C01873=-23.050,-43.100,93.800,0.0000,0.0000,-150.0000
C01874=-23.050,-38.100,93.800,0.0000,0.0000,-150.0000
C01875=-23.050,-33.100,93.800,0.0000,0.0000,-150.0000
C01876=-23.050,-28.100,93.800,0.0000,0.0000,-150.0000
C01877=-23.050,-23.100,93.800,0.0000,0.0000,-150.0000
C01878=-23.050,-18.100,93.800,0.0000,0.0000,-150.0000
C01879=-23.050,-13.100,93.800,0.0000,0.0000,-150.0000
C01880=-23.050,-8.100,93.800,0.0000,0.0000,-150.0000
C01881=-23.050,-3.100,93.800,0.0000,0.0000,-150.0000
C01882=-23.050,1.900,93.800,0.0000,0.0000,-150.0000
C01883=-23.050,6.900,93.800,0.0000,0.0000,-150.0000
C01884=-23.050,11.900,93.800,0.0000,0.0000,-150.0000
C01885=-23.050,16.900,93.800,0.0000,0.0000,-150.0000
C01886=-23.050,21.900,93.800,0.0000,0.0000,-150.0000
C01887=-23.050,26.900,93.800,0.0000,0.0000,-150.0000
C01888=-23.050,31.900,93.800,0.0000,0.0000,-150.0000
C01889=-23.050,36.900,93.800,0.0000,0.0000,-150.0000
C01890=-23.050,41.900,93.800,0.0000,0.0000,-150.0000
C01891=-18.267,41.900,93.800,0.0000,0.0000,-150.0000
C01892=-13.483,41.900,93.800,0.0000,0.0000,-150.0000
C01893=-8.700,41.900,93.800,0.0000,0.0000,-150.0000
C01894=-3.917,41.900,93.800,0.0000,0.0000,-150.0000
C01895=0.867,41.900,93.800,0.0000,0.0000,-150.0000
C01896=5.650,41.900,93.800,0.0000,0.0000,-150.0000
C01897=10.433,41.900,93.800,0.0000,0.0000,-150.0000
C01898=15.217,41.900,93.800,0.0000,0.0000,-150.0000
C01899=20.000,41.900,93.800,0.0000,0.0000,-150.0000
C01900=25.000,41.900,93.800,0.0000,0.0000,-150.0000
C01901=26.950,43.850,93.800,0.0000,0.0000,-150.0000
C01902=25.000,45.800,93.800,0.0000,0.0000,-150.0000
C01903=20.000,45.800,93.800,0.0000,0.0000,-150.0000
C01904=15.000,45.800,93.800,0.0000,0.0000,-150.0000
C01905=10.000,45.800,93.800,0.0000,0.0000,-150.0000
C01906=5.000,45.800,93.800,0.0000,0.0000,-150.0000
C01907=0.000,45.800,93.800,0.0000,0.0000,-150.0000
C01908=-5.000,45.800,93.800,0.0000,0.0000,-150.0000
C01909=-10.000,45.800,93.800,0.0000,0.0000,-150.0000
C01910=-15.000,45.800,93.800,0.0000,0.0000,-150.0000
C01911=-20.000,45.800,93.800,0.0000,0.0000,-150.0000
C01912=-25.000,45.800,93.800,0.0000,0.0000,-150.0000
C01913=-30.000,45.800,93.800,0.0000,0.0000,-150.0000
C01914=-35.000,45.800,93.800,0.0000,0.0000,-150.0000
C01915=-40.000,45.800,93.800,0.0000,0.0000,-150.0000
C01916=-45.000,45.800,93.800,0.0000,0.0000,-150.0000
C01917=-50.000,45.800,93.800,0.0000,0.0000,-150.0000
C01918=-55.000,45.800,93.800,0.0000,0.0000,-150.0000
C01919=-60.000,45.800,93.800,0.0000,0.0000,-150.0000
C01920=-65.000,45.800,93.800,0.0000,0.0000,-150.0000
C01921=-70.000,45.800,93.800,0.0000,0.0000,-150.0000
C01922=-75.000,45.800,93.800,0.0000,0.0000,-150.0000
C01923=-76.950,43.850,93.800,0.0000,0.0000,-150.0000
C01924=-75.000,41.900,93.800,0.0000,0.0000,-150.0000
C01925=-70.195,41.900,93.800,0.0000,0.0000,-150.0000
C01926=-65.390,41.900,93.800,0.0000,0.0000,-150.0000
C01927=-60.585,41.900,93.800,0.0000,0.0000,-150.0000
C01928=-55.780,41.900,93.800,0.0000,0.0000,-150.0000
C01929=-50.975,41.900,93.800,0.0000,0.0000,-150.0000
C01930=-46.170,41.900,93.800,0.0000,0.0000,-150.0000
C01931=-41.365,41.900,93.800,0.0000,0.0000,-150.0000
C01932=-36.560,41.900,93.800,0.0000,0.0000,-150.0000
C01933=-31.755,41.900,93.800,0.0000,0.0000,-150.0000
C01934=-26.950,41.900,93.800,0.0000,0.0000,-150.0000
C01935=-26.950,36.900,93.800,0.0000,0.0000,-150.0000
C01936=-26.950,31.900,93.800,0.0000,0.0000,-150.0000
C01937=-26.950,26.900,93.800,0.0000,0.0000,-150.0000
C01938=-26.950,21.900,93.800,0.0000,0.0000,-150.0000
C01939=-26.950,16.900,93.800,0.0000,0.0000,-150.0000
C01940=-26.950,11.900,93.800,0.0000,0.0000,-150.0000
C01941=-26.950,6.900,93.800,0.0000,0.0000,-150.0000
C01942=-26.950,1.900,93.800,0.0000,0.0000,-150.0000
C01943=-26.950,-3.100,93.800,0.0000,0.0000,-150.0000
C01944=-26.950,-8.100,93.800,0.0000,0.0000,-150.0000
C01945=-26.950,-13.100,93.800,0.0000,0.0000,-150.0000
C01946=-26.950,-18.100,93.800,0.0000,0.0000,-150.0000
C01947=-26.950,-23.100,93.800,0.0000,0.0000,-150.0000
C01948=-26.950,-28.100,93.800,0.0000,0.0000,-150.0000
C01949=-26.950,-33.100,93.800,0.0000,0.0000,-150.0000
C01950=-26.950,-38.100,93.800,0.0000,0.0000,-150.0000
C01951=-26.950,-43.100,93.800,0.0000,0.0000,-150.0000
C01952=-26.950,-48.100,93.800,0.0000,0.0000,-150.0000
C01953=-26.950,-53.100,93.800,0.0000,0.0000,-150.0000
C01954=-26.950,-58.100,93.800,0.0000,0.0000,-150.0000
C01955=-26.950,-63.100,93.800,0.0000,0.0000,-150.0000
C01956=-26.950,-68.100,93.800,0.0000,0.0000,-150.0000
C01957=-31.755,-68.100,93.800,0.0000,0.0000,-150.0000
C01958=-36.560,-68.100,93.800,0.0000,0.0000,-150.0000
C01959=-41.365,-68.100,93.800,0.0000,0.0000,-150.0000
C01960=-46.170,-68.100,93.800,0.0000,0.0000,-150.0000
C01961=-50.975,-68.100,93.800,0.0000,0.0000,-150.0000
C01962=-55.780,-68.100,93.800,0.0000,0.0000,-150.0000
C01963=-60.585,-68.100,93.800,0.0000,0.0000,-150.0000
C01964=-65.390,-68.100,93.800,0.0000,0.0000,-150.0000
C01965=-70.195,-68.100,93.800,0.0000,0.0000,-150.0000
C01966=-75.000,-68.100,93.800,0.0000,0.0000,-150.0000
C01967=-75.000,-68.100,95.500,0.0000,0.0000,-150.0000
C01968=-70.195,-68.100,95.500,0.0000,0.0000,-150.0000
C01969=-65.390,-68.100,95.500,0.0000,0.0000,-150.0000
C01970=-60.585,-68.100,95.500,0.0000,0.0000,-150.0000
C01971=-55.780,-68.100,95.500,0.0000,0.0000,-150.0000
C01972=-50.975,-68.100,95.500,0.0000,0.0000,-150.0000
C01973=-46.170,-68.100,95.500,0.0000,0.0000,-150.0000
C01974=-41.365,-68.100,95.500,0.0000,0.0000,-150.0000
C01975=-36.560,-68.100,95.500,0.0000,0.0000,-150.0000
C01976=-31.755,-68.100,95.500,0.0000,0.0000,-150.0000
C01977=-26.950,-68.100,95.500,0.0000,0.0000,-150.0000
C01978=-26.950,-63.100,95.500,0.0000,0.0000,-150.0000
C01979=-26.950,-58.100,95.500,0.0000,0.0000,-150.0000
C01980=-26.950,-53.100,95.500,0.0000,0.0000,-150.0000
C01981=-26.950,-48.100,95.500,0.0000,0.0000,-150.0000
C01982=-26.950,-43.100,95.500,0.0000,0.0000,-150.0000
C01983=-26.950,-38.100,95.500,0.0000,0.0000,-150.0000
C01984=-26.950,-33.100,95.500,0.0000,0.0000,-150.0000
C01985=-26.950,-28.100,95.500,0.0000,0.0000,-150.0000
C01986=-26.950,-23.100,95.500,0.0000,0.0000,-150.0000
C01987=-26.950,-18.100,95.500,0.0000,0.0000,-150.0000
C01988=-26.950,-13.100,95.500,0.0000,0.0000,-150.0000
C01989=-26.950,-8.100,95.500,0.0000,0.0000,-150.0000
C01990=-26.950,-3.100,95.500,0.0000,0.0000,-150.0000
C01991=-26.950,1.900,95.500,0.0000,0.0000,-150.0000
C01992=-26.950,6.900,95.500,0.0000,0.0000,-150.0000
C01993=-26.950,11.900,95.500,0.0000,0.0000,-150.0000
C01994=-26.950,16.900,95.500,0.0000,0.0000,-150.0000
C01995=-26.950,21.900,95.500,0.0000,0.0000,-150.0000
C01996=-26.950,26.900,95.500,0.0000,0.0000,-150.0000
C01997=-26.950,31.900,95.500,0.0000,0.0000,-150.0000
C01998=-26.950,36.900,95.500,0.0000,0.0000,-150.0000
C01999=-26.950,41.900,95.500,0.0000,0.0000,-150.0000
C02000=-31.733,41.900,95.500,0.0000,0.0000,-150.0000
C02001=-36.517,41.900,95.500,0.0000,0.0000,-150.0000
C02002=-41.300,41.900,95.500,0.0000,0.0000,-150.0000
C02003=-46.083,41.900,95.500,0.0000,0.0000,-150.0000
C02004=-50.867,41.900,95.500,0.0000,0.0000,-150.0000
C02005=-55.650,41.900,95.500,0.0000,0.0000,-150.0000
C02006=-60.433,41.900,95.500,0.0000,0.0000,-150.0000
C02007=-65.217,41.900,95.500,0.0000,0.0000,-150.0000
C02008=-70.000,41.900,95.500,0.0000,0.0000,-150.0000
C02009=-75.000,41.900,95.500,0.0000,0.0000,-150.0000
C02010=-76.950,43.850,95.500,0.0000,0.0000,-150.0000
C02011=-75.000,45.800,95.500,0.0000,0.0000,-150.0000
C02012=-70.000,45.800,95.500,0.0000,0.0000,-150.0000
C02013=-65.000,45.800,95.500,0.0000,0.0000,-150.0000
C02014=-60.000,45.800,95.500,0.0000,0.0000,-150.0000
C02015=-55.000,45.800,95.500,0.0000,0.0000,-150.0000
C02016=-50.000,45.800,95.500,0.0000,0.0000,-150.0000
C02017=-45.000,45.800,95.500,0.0000,0.0000,-150.0000
C02018=-40.000,45.800,95.500,0.0000,0.0000,-150.0000
C02019=-35.000,45.800,95.500,0.0000,0.0000,-150.0000
C02020=-30.000,45.800,95.500,0.0000,0.0000,-150.0000
C02021=-25.000,45.800,95.500,0.0000,0.0000,-150.0000
C02022=-20.000,45.800,95.500,0.0000,0.0000,-150.0000
C02023=-15.000,45.800,95.500,0.0000,0.0000,-150.0000
C02024=-10.000,45.800,95.500,0.0000,0.0000,-150.0000
C02025=-5.000,45.800,95.500,0.0000,0.0000,-150.0000
C02026=0.000,45.800,95.500,0.0000,0.0000,-150.0000
C02027=5.000,45.800,95.500,0.0000,0.0000,-150.0000
C02028=10.000,45.800,95.500,0.0000,0.0000,-150.0000
C02029=15.000,45.800,95.500,0.0000,0.0000,-150.0000
C02030=20.000,45.800,95.500,0.0000,0.0000,-150.0000
C02031=25.000,45.800,95.500,0.0000,0.0000,-150.0000
C02032=26.950,43.850,95.500,0.0000,0.0000,-150.0000
C02033=25.000,41.900,95.500,0.0000,0.0000,-150.0000
C02034=20.195,41.900,95.500,0.0000,0.0000,-150.0000
C02035=15.390,41.900,95.500,0.0000,0.0000,-150.0000
C02036=10.585,41.900,95.500,0.0000,0.0000,-150.0000
C02037=5.780,41.900,95.500,0.0000,0.0000,-150.0000
C02038=0.975,41.900,95.500,0.0000,0.0000,-150.0000
C02039=-3.830,41.900,95.500,0.0000,0.0000,-150.0000
C02040=-8.635,41.900,95.500,0.0000,0.0000,-150.0000
C02041=-13.440,41.900,95.500,0.0000,0.0000,-150.0000
C02042=-18.245,41.900,95.500,0.0000,0.0000,-150.0000
C02043=-23.050,41.900,95.500,0.0000,0.0000,-150.0000
C02044=-23.050,36.900,95.500,0.0000,0.0000,-150.0000
C02045=-23.050,31.900,95.500,0.0000,0.0000,-150.0000
C02046=-23.050,26.900,95.500,0.0000,0.0000,-150.0000
C02047=-23.050,21.900,95.500,0.0000,0.0000,-150.0000
C02048=-23.050,16.900,95.500,0.0000,0.0000,-150.0000
C02049=-23.050,11.900,95.500,0.0000,0.0000,-150.0000
C02050=-23.050,6.900,95.500,0.0000,0.0000,-150.0000
C02051=-23.050,1.900,95.500,0.0000,0.0000,-150.0000
C02052=-23.050,-3.100,95.500,0.0000,0.0000,-150.0000
C02053=-23.050,-8.100,95.500,0.0000,0.0000,-150.0000
C02054=-23.050,-13.100,95.500,0.0000,0.0000,-150.0000
C02055=-23.050,-18.100,95.500,0.0000,0.0000,-150.0000
C02056=-23.050,-23.100,95.500,0.0000,0.0000,-150.0000
C02057=-23.050,-28.100,95.500,0.0000,0.0000,-150.0000
C02058=-23.050,-33.100,95.500,0.0000,0.0000,-150.0000
C02059=-23.050,-38.100,95.500,0.0000,0.0000,-150.0000
C02060=-23.050,-43.100,95.500,0.0000,0.0000,-150.0000
C02061=-23.050,-48.100,95.500,0.0000,0.0000,-150.0000
C02062=-23.050,-53.100,95.500,0.0000,0.0000,-150.0000
C02063=-23.050,-58.100,95.500,0.0000,0.0000,-150.0000
C02064=-23.050,-63.100,95.500,0.0000,0.0000,-150.0000
C02065=-23.050,-68.100,95.500,0.0000,0.0000,-150.0000
C02066=-18.267,-68.100,95.500,0.0000,0.0000,-150.0000
C02067=-13.483,-68.100,95.500,0.0000,0.0000,-150.0000
C02068=-8.700,-68.100,95.500,0.0000,0.0000,-150.0000
C02069=-3.917,-68.100,95.500,0.0000,0.0000,-150.0000
C02070=0.867,-68.100,95.500,0.0000,0.0000,-150.0000
C02071=5.650,-68.100,95.500,0.0000,0.0000,-150.0000
C02072=10.433,-68.100,95.500,0.0000,0.0000,-150.0000
C02073=15.217,-68.100,95.500,0.0000,0.0000,-150.0000
C02074=20.000,-68.100,95.500,0.0000,0.0000,-150.0000
C02075=25.000,-68.100,95.500,0.0000,0.0000,-150.0000
C02076=26.950,-70.050,95.500,0.0000,0.0000,-150.0000
C02077=25.000,-72.000,95.500,0.0000,0.0000,-150.0000
C02078=20.000,-72.000,95.500,0.0000,0.0000,-150.0000
C02079=15.000,-72.000,95.500,0.0000,0.0000,-150.0000
C02080=10.000,-72.000,95.500,0.0000,0.0000,-150.0000
C02081=5.000,-72.000,95.500,0.0000,0.0000,-150.0000
C02082=0.000,-72.000,95.500,0.0000,0.0000,-150.0000
C02083=-5.000,-72.000,95.500,0.0000,0.0000,-150.0000
C02084=-10.000,-72.000,95.500,0.0000,0.0000,-150.0000
C02085=-15.000,-72.000,95.500,0.0000,0.0000,-150.0000
C02086=-20.000,-72.000,95.500,0.0000,0.0000,-150.0000
C02087=-25.000,-72.000,95.500,0.0000,0.0000,-150.0000
C02088=-30.000,-72.000,95.500,0.0000,0.0000,-150.0000
C02089=-35.000,-72.000,95.500,0.0000,0.0000,-150.0000
C02090=-40.000,-72.000,95.500,0.0000,0.0000,-150.0000
C02091=-45.000,-72.000,95.500,0.0000,0.0000,-150.0000
C02092=-50.000,-72.000,95.500,0.0000,0.0000,-150.0000
C02093=-55.000,-72.000,95.500,0.0000,0.0000,-150.0000
C02094=-60.000,-72.000,95.500,0.0000,0.0000,-150.0000
C02095=-65.000,-72.000,95.500,0.0000,0.0000,-150.0000
C02096=-70.000,-72.000,95.500,0.0000,0.0000,-150.0000
C02097=-75.000,-72.000,95.500,0.0000,0.0000,-150.0000
C02098=-75.000,-72.000,97.200,0.0000,0.0000,-150.0000
C02099=-70.000,-72.000,97.200,0.0000,0.0000,-150.0000
C02100=-65.000,-72.000,97.200,0.0000,0.0000,-150.0000
C02101=-60.000,-72.000,97.200,0.0000,0.0000,-150.0000
C02102=-55.000,-72.000,97.200,0.0000,0.0000,-150.0000
C02103=-50.000,-72.000,97.200,0.0000,0.0000,-150.0000
C02104=-45.000,-72.000,97.200,0.0000,0.0000,-150.0000
C02105=-40.000,-72.000,97.200,0.0000,0.0000,-150.0000
C02106=-35.000,-72.000,97.200,0.0000,0.0000,-150.0000
C02107=-30.000,-72.000,97.200,0.0000,0.0000,-150.0000
C02108=-25.000,-72.000,97.200,0.0000,0.0000,-150.0000
C02109=-20.000,-72.000,97.200,0.0000,0.0000,-150.0000
C02110=-15.000,-72.000,97.200,0.0000,0.0000,-150.0000
C02111=-10.000,-72.000,97.200,0.0000,0.0000,-150.0000
C02112=-5.000,-72.000,97.200,0.0000,0.0000,-150.0000
C02113=0.000,-72.000,97.200,0.0000,0.0000,-150.0000
C02114=5.000,-72.000,97.200,0.0000,0.0000,-150.0000
C02115=10.000,-72.000,97.200,0.0000,0.0000,-150.0000
C02116=15.000,-72.000,97.200,0.0000,0.0000,-150.0000
C02117=20.000,-72.000,97.200,0.0000,0.0000,-150.0000
C02118=25.000,-72.000,97.200,0.0000,0.0000,-150.0000
C02119=26.950,-70.050,97.200,0.0000,0.0000,-150.0000
C02120=25.000,-68.100,97.200,0.0000,0.0000,-150.0000
C02121=20.195,-68.100,97.200,0.0000,0.0000,-150.0000
C02122=15.390,-68.100,97.200,0.0000,0.0000,-150.0000
C02123=10.585,-68.100,97.200,0.0000,0.0000,-150.0000
C02124=5.780,-68.100,97.200,0.0000,0.0000,-150.0000
C02125=0.975,-68.100,97.200,0.0000,0.0000,-150.0000
C02126=-3.830,-68.100,97.200,0.0000,0.0000,-150.0000
C02127=-8.635,-68.100,97.200,0.0000,0.0000,-150.0000
C02128=-13.440,-68.100,97.200,0.0000,0.0000,-150.0000
C02129=-18.245,-68.100,97.200,0.0000,0.0000,-150.0000
C02130=-23.050,-68.100,97.200,0.0000,0.0000,-150.0000
C02131=-23.050,-63.100,97.200,0.0000,0.0000,-150.0000
C02132=-23.050,-58.100,97.200,0.0000,0.0000,-150.0000
C02133=-23.050,-53.100,97.200,0.0000,0.0000,-150.0000
C02134=-23.050,-48.100,97.200,0.0000,0.0000,-150.0000
C02135=-23.050,-43.100,97.200,0.0000,0.0000,-150.0000
C02136=-23.050,-38.100,97.200,0.0000,0.0000,-150.0000
C02137=-23.050,-33.100,97.200,0.0000,0.0000,-150.0000
C02138=-23.050,-28.100,97.200,0.0000,0.0000,-150.0000
C02139=-23.050,-23.100,97.200,0.0000,0.0000,-150.0000
C02140=-23.050,-18.100,97.200,0.0000,0.0000,-150.0000
C02141=-23.050,-13.100,97.200,0.0000,0.0000,-150.0000
C02142=-23.050,-8.100,97.200,0.0000,0.0000,-150.0000
C02143=-23.050,-3.100,97.200,0.0000,0.0000,-150.0000
C02144=-23.050,1.900,97.200,0.0000,0.0000,-150.0000
C02145=-23.050,6.900,97.200,0.0000,0.0000,-150.0000
C02146=-23.050,11.900,97.200,0.0000,0.0000,-150.0000
C02147=-23.050,16.900,97.200,0.0000,0.0000,-150.0000
C02148=-23.050,21.900,97.200,0.0000,0.0000,-150.0000
C02149=-23.050,26.900,97.200,0.0000,0.0000,-150.0000
C02150=-23.050,31.900,97.200,0.0000,0.0000,-150.0000
C02151=-23.050,36.900,97.200,0.0000,0.0000,-150.0000
C02152=-23.050,41.900,97.200,0.0000,0.0000,-150.0000
C02153=-18.267,41.900,97.200,0.0000,0.0000,-150.0000
C02154=-13.483,41.900,97.200,0.0000,0.0000,-150.0000
C02155=-8.700,41.900,97.200,0.0000,0.0000,-150.0000
C02156=-3.917,41.900,97.200,0.0000,0.0000,-150.0000
C02157=0.867,41.900,97.200,0.0000,0.0000,-150.0000
C02158=5.650,41.900,97.200,0.0000,0.0000,-150.0000
C02159=10.433,41.900,97.200,0.0000,0.0000,-150.0000
C02160=15.217,41.900,97.200,0.0000,0.0000,-150.0000
C02161=20.000,41.900,97.200,0.0000,0.0000,-150.0000
C02162=25.000,41.900,97.200,0.0000,0.0000,-150.0000
C02163=26.950,43.850,97.200,0.0000,0.0000,-150.0000
C02164=25.000,45.800,97.200,0.0000,0.0000,-150.0000
C02165=20.000,45.800,97.200,0.0000,0.0000,-150.0000
C02166=15.000,45.800,97.200,0.0000,0.0000,-150.0000
C02167=10.000,45.800,97.200,0.0000,0.0000,-150.0000
C02168=5.000,45.800,97.200,0.0000,0.0000,-150.0000
C02169=0.000,45.800,97.200,0.0000,0.0000,-150.0000
C02170=-5.000,45.800,97.200,0.0000,0.0000,-150.0000
C02171=-10.000,45.800,97.200,0.0000,0.0000,-150.0000
C02172=-15.000,45.800,97.200,0.0000,0.0000,-150.0000
C02173=-20.000,45.800,97.200,0.0000,0.0000,-150.0000
C02174=-25.000,45.800,97.200,0.0000,0.0000,-150.0000
C02175=-30.000,45.800,97.200,0.0000,0.0000,-150.0000
C02176=-35.000,45.800,97.200,0.0000,0.0000,-150.0000
C02177=-40.000,45.800,97.200,0.0000,0.0000,-150.0000
C02178=-45.000,45.800,97.200,0.0000,0.0000,-150.0000
C02179=-50.000,45.800,97.200,0.0000,0.0000,-150.0000
C02180=-55.000,45.800,97.200,0.0000,0.0000,-150.0000
C02181=-60.000,45.800,97.200,0.0000,0.0000,-150.0000
C02182=-65.000,45.800,97.200,0.0000,0.0000,-150.0000
C02183=-70.000,45.800,97.200,0.0000,0.0000,-150.0000
C02184=-75.000,45.800,97.200,0.0000,0.0000,-150.0000
C02185=-76.950,43.850,97.200,0.0000,0.0000,-150.0000
C02186=-75.000,41.900,97.200,0.0000,0.0000,-150.0000
C02187=-70.195,41.900,97.200,0.0000,0.0000,-150.0000
C02188=-65.390,41.900,97.200,0.0000,0.0000,-150.0000
C02189=-60.585,41.900,97.200,0.0000,0.0000,-150.0000
C02190=-55.780,41.900,97.200,0.0000,0.0000,-150.0000
C02191=-50.975,41.900,97.200,0.0000,0.0000,-150.0000
C02192=-46.170,41.900,97.200,0.0000,0.0000,-150.0000
C02193=-41.365,41.900,97.200,0.0000,0.0000,-150.0000
C02194=-36.560,41.900,97.200,0.0000,0.0000,-150.0000
C02195=-31.755,41.900,97.200,0.0000,0.0000,-150.0000
C02196=-26.950,41.900,97.200,0.0000,0.0000,-150.0000
C02197=-26.950,36.900,97.200,0.0000,0.0000,-150.0000
C02198=-26.950,31.900,97.200,0.0000,0.0000,-150.0000
C02199=-26.950,26.900,97.200,0.0000,0.0000,-150.0000
C02200=-26.950,21.900,97.200,0.0000,0.0000,-150.0000
C02201=-26.950,16.900,97.200,0.0000,0.0000,-150.0000
C02202=-26.950,11.900,97.200,0.0000,0.0000,-150.0000
C02203=-26.950,6.900,97.200,0.0000,0.0000,-150.0000
C02204=-26.950,1.900,97.200,0.0000,0.0000,-150.0000
C02205=-26.950,-3.100,97.200,0.0000,0.0000,-150.0000
C02206=-26.950,-8.100,97.200,0.0000,0.0000,-150.0000
C02207=-26.950,-13.100,97.200,0.0000,0.0000,-150.0000
C02208=-26.950,-18.100,97.200,0.0000,0.0000,-150.0000
C02209=-26.950,-23.100,97.200,0.0000,0.0000,-150.0000
C02210=-26.950,-28.100,97.200,0.0000,0.0000,-150.0000
C02211=-26.950,-33.100,97.200,0.0000,0.0000,-150.0000
C02212=-26.950,-38.100,97.200,0.0000,0.0000,-150.0000
C02213=-26.950,-43.100,97.200,0.0000,0.0000,-150.0000
C02214=-26.950,-48.100,97.200,0.0000,0.0000,-150.0000
C02215=-26.950,-53.100,97.200,0.0000,0.0000,-150.0000
C02216=-26.950,-58.100,97.200,0.0000,0.0000,-150.0000
C02217=-26.950,-63.100,97.200,0.0000,0.0000,-150.0000
C02218=-26.950,-68.100,97.200,0.0000,0.0000,-150.0000
C02219=-31.755,-68.100,97.200,0.0000,0.0000,-150.0000
C02220=-36.560,-68.100,97.200,0.0000,0.0000,-150.0000
C02221=-41.365,-68.100,97.200,0.0000,0.0000,-150.0000
C02222=-46.170,-68.100,97.200,0.0000,0.0000,-150.0000
C02223=-50.975,-68.100,97.200,0.0000,0.0000,-150.0000
C02224=-55.780,-68.100,97.200,0.0000,0.0000,-150.0000
C02225=-60.585,-68.100,97.200,0.0000,0.0000,-150.0000
C02226=-65.390,-68.100,97.200,0.0000,0.0000,-150.0000
C02227=-70.195,-68.100,97.200,0.0000,0.0000,-150.0000
C02228=-75.000,-68.100,97.200,0.0000,0.0000,-150.0000
C02229=-75.000,-68.100,98.900,0.0000,0.0000,-150.0000
C02230=-70.195,-68.100,98.900,0.0000,0.0000,-150.0000
C02231=-65.390,-68.100,98.900,0.0000,0.0000,-150.0000
C02232=-60.585,-68.100,98.900,0.0000,0.0000,-150.0000
C02233=-55.780,-68.100,98.900,0.0000,0.0000,-150.0000
C02234=-50.975,-68.100,98.900,0.0000,0.0000,-150.0000
C02235=-46.170,-68.100,98.900,0.0000,0.0000,-150.0000
C02236=-41.365,-68.100,98.900,0.0000,0.0000,-150.0000
C02237=-36.560,-68.100,98.900,0.0000,0.0000,-150.0000
C02238=-31.755,-68.100,98.900,0.0000,0.0000,-150.0000
C02239=-26.950,-68.100,98.900,0.0000,0.0000,-150.0000
C02240=-26.950,-63.100,98.900,0.0000,0.0000,-150.0000
C02241=-26.950,-58.100,98.900,0.0000,0.0000,-150.0000
C02242=-26.950,-53.100,98.900,0.0000,0.0000,-150.0000
C02243=-26.950,-48.100,98.900,0.0000,0.0000,-150.0000
C02244=-26.950,-43.100,98.900,0.0000,0.0000,-150.0000
C02245=-26.950,-38.100,98.900,0.0000,0.0000,-150.0000
C02246=-26.950,-33.100,98.900,0.0000,0.0000,-150.0000
C02247=-26.950,-28.100,98.900,0.0000,0.0000,-150.0000
C02248=-26.950,-23.100,98.900,0.0000,0.0000,-150.0000
C02249=-26.950,-18.100,98.900,0.0000,0.0000,-150.0000
C02250=-26.950,-13.100,98.900,0.0000,0.0000,-150.0000
C02251=-26.950,-8.100,98.900,0.0000,0.0000,-150.0000
C02252=-26.950,-3.100,98.900,0.0000,0.0000,-150.0000
C02253=-26.950,1.900,98.900,0.0000,0.0000,-150.0000
C02254=-26.950,6.900,98.900,0.0000,0.0000,-150.0000
C02255=-26.950,11.900,98.900,0.0000,0.0000,-150.0000
C02256=-26.950,16.900,98.900,0.0000,0.0000,-150.0000
C02257=-26.950,21.900,98.900,0.0000,0.0000,-150.0000
C02258=-26.950,26.900,98.900,0.0000,0.0000,-150.0000
C02259=-26.950,31.900,98.900,0.0000,0.0000,-150.0000
C02260=-26.950,36.900,98.900,0.0000,0.0000,-150.0000
C02261=-26.950,41.900,98.900,0.0000,0.0000,-150.0000
C02262=-31.733,41.900,98.900,0.0000,0.0000,-150.0000
C02263=-36.517,41.900,98.900,0.0000,0.0000,-150.0000
C02264=-41.300,41.900,98.900,0.0000,0.0000,-150.0000
C02265=-46.083,41.900,98.900,0.0000,0.0000,-150.0000
C02266=-50.867,41.900,98.900,0.0000,0.0000,-150.0000
C02267=-55.650,41.900,98.900,0.0000,0.0000,-150.0000
C02268=-60.433,41.900,98.900,0.0000,0.0000,-150.0000
C02269=-65.217,41.900,98.900,0.0000,0.0000,-150.0000
C02270=-70.000,41.900,98.900,0.0000,0.0000,-150.0000
C02271=-75.000,41.900,98.900,0.0000,0.0000,-150.0000
C02272=-76.950,43.850,98.900,0.0000,0.0000,-150.0000
C02273=-75.000,45.800,98.900,0.0000,0.0000,-150.0000
C02274=-70.000,45.800,98.900,0.0000,0.0000,-150.0000
C02275=-65.000,45.800,98.900,0.0000,0.0000,-150.0000
C02276=-60.000,45.800,98.900,0.0000,0.0000,-150.0000
C02277=-55.000,45.800,98.900,0.0000,0.0000,-150.0000
C02278=-50.000,45.800,98.900,0.0000,0.0000,-150.0000
C02279=-45.000,45.800,98.900,0.0000,0.0000,-150.0000
C02280=-40.000,45.800,98.900,0.0000,0.0000,-150.0000
C02281=-35.000,45.800,98.900,0.0000,0.0000,-150.0000
C02282=-30.000,45.800,98.900,0.0000,0.0000,-150.0000
C02283=-25.000,45.800,98.900,0.0000,0.0000,-150.0000
C02284=-20.000,45.800,98.900,0.0000,0.0000,-150.0000
C02285=-15.000,45.800,98.900,0.0000,0.0000,-150.0000
C02286=-10.000,45.800,98.900,0.0000,0.0000,-150.0000
C02287=-5.000,45.800,98.900,0.0000,0.0000,-150.0000
C02288=0.000,45.800,98.900,0.0000,0.0000,-150.0000
C02289=5.000,45.800,98.900,0.0000,0.0000,-150.0000
C02290=10.000,45.800,98.900,0.0000,0.0000,-150.0000
C02291=15.000,45.800,98.900,0.0000,0.0000,-150.0000
C02292=20.000,45.800,98.900,0.0000,0.0000,-150.0000
C02293=25.000,45.800,98.900,0.0000,0.0000,-150.0000
C02294=26.950,43.850,98.900,0.0000,0.0000,-150.0000
C02295=25.000,41.900,98.900,0.0000,0.0000,-150.0000
C02296=20.195,41.900,98.900,0.0000,0.0000,-150.0000
C02297=15.390,41.900,98.900,0.0000,0.0000,-150.0000
C02298=10.585,41.900,98.900,0.0000,0.0000,-150.0000
C02299=5.780,41.900,98.900,0.0000,0.0000,-150.0000
C02300=0.975,41.900,98.900,0.0000,0.0000,-150.0000
C02301=-3.830,41.900,98.900,0.0000,0.0000,-150.0000
C02302=-8.635,41.900,98.900,0.0000,0.0000,-150.0000
C02303=-13.440,41.900,98.900,0.0000,0.0000,-150.0000
C02304=-18.245,41.900,98.900,0.0000,0.0000,-150.0000
C02305=-23.050,41.900,98.900,0.0000,0.0000,-150.0000
C02306=-23.050,36.900,98.900,0.0000,0.0000,-150.0000
C02307=-23.050,31.900,98.900,0.0000,0.0000,-150.0000
C02308=-23.050,26.900,98.900,0.0000,0.0000,-150.0000
C02309=-23.050,21.900,98.900,0.0000,0.0000,-150.0000
C02310=-23.050,16.900,98.900,0.0000,0.0000,-150.0000
C02311=-23.050,11.900,98.900,0.0000,0.0000,-150.0000
C02312=-23.050,6.900,98.900,0.0000,0.0000,-150.0000
C02313=-23.050,1.900,98.900,0.0000,0.0000,-150.0000
C02314=-23.050,-3.100,98.900,0.0000,0.0000,-150.0000
C02315=-23.050,-8.100,98.900,0.0000,0.0000,-150.0000
C02316=-23.050,-13.100,98.900,0.0000,0.0000,-150.0000
C02317=-23.050,-18.100,98.900,0.0000,0.0000,-150.0000
C02318=-23.050,-23.100,98.900,0.0000,0.0000,-150.0000
C02319=-23.050,-28.100,98.900,0.0000,0.0000,-150.0000
C02320=-23.050,-33.100,98.900,0.0000,0.0000,-150.0000
C02321=-23.050,-38.100,98.900,0.0000,0.0000,-150.0000
C02322=-23.050,-43.100,98.900,0.0000,0.0000,-150.0000
C02323=-23.050,-48.100,98.900,0.0000,0.0000,-150.0000
C02324=-23.050,-53.100,98.900,0.0000,0.0000,-150.0000
C02325=-23.050,-58.100,98.900,0.0000,0.0000,-150.0000
C02326=-23.050,-63.100,98.900,0.0000,0.0000,-150.0000
C02327=-23.050,-68.100,98.900,0.0000,0.0000,-150.0000
C02328=-18.267,-68.100,98.900,0.0000,0.0000,-150.0000
C02329=-13.483,-68.100,98.900,0.0000,0.0000,-150.0000
C02330=-8.700,-68.100,98.900,0.0000,0.0000,-150.0000
C02331=-3.917,-68.100,98.900,0.0000,0.0000,-150.0000
C02332=0.867,-68.100,98.900,0.0000,0.0000,-150.0000
C02333=5.650,-68.100,98.900,0.0000,0.0000,-150.0000
C02334=10.433,-68.100,98.900,0.0000,0.0000,-150.0000
C02335=15.217,-68.100,98.900,0.0000,0.0000,-150.0000
C02336=20.000,-68.100,98.900,0.0000,0.0000,-150.0000
C02337=25.000,-68.100,98.900,0.0000,0.0000,-150.0000
C02338=26.950,-70.050,98.900,0.0000,0.0000,-150.0000
C02339=25.000,-72.000,98.900,0.0000,0.0000,-150.0000
C02340=20.000,-72.000,98.900,0.0000,0.0000,-150.0000
C02341=15.000,-72.000,98.900,0.0000,0.0000,-150.0000
C02342=10.000,-72.000,98.900,0.0000,0.0000,-150.0000
C02343=5.000,-72.000,98.900,0.0000,0.0000,-150.0000
C02344=0.000,-72.000,98.900,0.0000,0.0000,-150.0000
C02345=-5.000,-72.000,98.900,0.0000,0.0000,-150.0000
C02346=-10.000,-72.000,98.900,0.0000,0.0000,-150.0000
C02347=-15.000,-72.000,98.900,0.0000,0.0000,-150.0000
C02348=-20.000,-72.000,98.900,0.0000,0.0000,-150.0000
C02349=-25.000,-72.000,98.900,0.0000,0.0000,-150.0000
C02350=-30.000,-72.000,98.900,0.0000,0.0000,-150.0000
C02351=-35.000,-72.000,98.900,0.0000,0.0000,-150.0000
C02352=-40.000,-72.000,98.900,0.0000,0.0000,-150.0000
C02353=-45.000,-72.000,98.900,0.0000,0.0000,-150.0000
C02354=-50.000,-72.000,98.900,0.0000,0.0000,-150.0000
C02355=-55.000,-72.000,98.900,0.0000,0.0000,-150.0000
C02356=-60.000,-72.000,98.900,0.0000,0.0000,-150.0000
C02357=-65.000,-72.000,98.900,0.0000,0.0000,-150.0000
C02358=-70.000,-72.000,98.900,0.0000,0.0000,-150.0000
C02359=-75.000,-72.000,98.900,0.0000,0.0000,-150.0000
C02360=-75.000,-72.000,100.600,0.0000,0.0000,-150.0000
C02361=-70.000,-72.000,100.600,0.0000,0.0000,-150.0000
C02362=-65.000,-72.000,100.600,0.0000,0.0000,-150.0000
C02363=-60.000,-72.000,100.600,0.0000,0.0000,-150.0000
C02364=-55.000,-72.000,100.600,0.0000,0.0000,-150.0000
C02365=-50.000,-72.000,100.600,0.0000,0.0000,-150.0000
C02366=-45.000,-72.000,100.600,0.0000,0.0000,-150.0000
C02367=-40.000,-72.000,100.600,0.0000,0.0000,-150.0000
C02368=-35.000,-72.000,100.600,0.0000,0.0000,-150.0000
C02369=-30.000,-72.000,100.600,0.0000,0.0000,-150.0000
C02370=-25.000,-72.000,100.600,0.0000,0.0000,-150.0000
C02371=-20.000,-72.000,100.600,0.0000,0.0000,-150.0000
C02372=-15.000,-72.000,100.600,0.0000,0.0000,-150.0000
C02373=-10.000,-72.000,100.600,0.0000,0.0000,-150.0000
C02374=-5.000,-72.000,100.600,0.0000,0.0000,-150.0000
C02375=0.000,-72.000,100.600,0.0000,0.0000,-150.0000
C02376=5.000,-72.000,100.600,0.0000,0.0000,-150.0000
C02377=10.000,-72.000,100.600,0.0000,0.0000,-150.0000
C02378=15.000,-72.000,100.600,0.0000,0.0000,-150.0000
C02379=20.000,-72.000,100.600,0.0000,0.0000,-150.0000
C02380=25.000,-72.000,100.600,0.0000,0.0000,-150.0000
C02381=26.950,-70.050,100.600,0.0000,0.0000,-150.0000
C02382=25.000,-68.100,100.600,0.0000,0.0000,-150.0000
C02383=20.195,-68.100,100.600,0.0000,0.0000,-150.0000
C02384=15.390,-68.100,100.600,0.0000,0.0000,-150.0000
C02385=10.585,-68.100,100.600,0.0000,0.0000,-150.0000
C02386=5.780,-68.100,100.600,0.0000,0.0000,-150.0000
C02387=0.975,-68.100,100.600,0.0000,0.0000,-150.0000
C02388=-3.830,-68.100,100.600,0.0000,0.0000,-150.0000
C02389=-8.635,-68.100,100.600,0.0000,0.0000,-150.0000
C02390=-13.440,-68.100,100.600,0.0000,0.0000,-150.0000
C02391=-18.245,-68.100,100.600,0.0000,0.0000,-150.0000
C02392=-23.050,-68.100,100.600,0.0000,0.0000,-150.0000
C02393=-23.050,-63.100,100.600,0.0000,0.0000,-150.0000
C02394=-23.050,-58.100,100.600,0.0000,0.0000,-150.0000
C02395=-23.050,-53.100,100.600,0.0000,0.0000,-150.0000
C02396=-23.050,-48.100,100.600,0.0000,0.0000,-150.0000
C02397=-23.050,-43.100,100.600,0.0000,0.0000,-150.0000
C02398=-23.050,-38.100,100.600,0.0000,0.0000,-150.0000
C02399=-23.050,-33.100,100.600,0.0000,0.0000,-150.0000
C02400=-23.050,-28.100,100.600,0.0000,0.0000,-150.0000
C02401=-23.050,-23.100,100.600,0.0000,0.0000,-150.0000
C02402=-23.050,-18.100,100.600,0.0000,0.0000,-150.0000
C02403=-23.050,-13.100,100.600,0.0000,0.0000,-150.0000
C02404=-23.050,-8.100,100.600,0.0000,0.0000,-150.0000
C02405=-23.050,-3.100,100.600,0.0000,0.0000,-150.0000
C02406=-23.050,1.900,100.600,0.0000,0.0000,-150.0000
C02407=-23.050,6.900,100.600,0.0000,0.0000,-150.0000
C02408=-23.050,11.900,100.600,0.0000,0.0000,-150.0000
C02409=-23.050,16.900,100.600,0.0000,0.0000,-150.0000
C02410=-23.050,21.900,100.600,0.0000,0.0000,-150.0000
C02411=-23.050,26.900,100.600,0.0000,0.0000,-150.0000
C02412=-23.050,31.900,100.600,0.0000,0.0000,-150.0000
C02413=-23.050,36.900,100.600,0.0000,0.0000,-150.0000
C02414=-23.050,41.900,100.600,0.0000,0.0000,-150.0000
C02415=-18.267,41.900,100.600,0.0000,0.0000,-150.0000
C02416=-13.483,41.900,100.600,0.0000,0.0000,-150.0000
C02417=-8.700,41.900,100.600,0.0000,0.0000,-150.0000
C02418=-3.917,41.900,100.600,0.0000,0.0000,-150.0000
C02419=0.867,41.900,100.600,0.0000,0.0000,-150.0000
C02420=5.650,41.900,100.600,0.0000,0.0000,-150.0000
C02421=10.433,41.900,100.600,0.0000,0.0000,-150.0000
C02422=15.217,41.900,100.600,0.0000,0.0000,-150.0000
C02423=20.000,41.900,100.600,0.0000,0.0000,-150.0000
C02424=25.000,41.900,100.600,0.0000,0.0000,-150.0000
C02425=26.950,43.850,100.600,0.0000,0.0000,-150.0000
C02426=25.000,45.800,100.600,0.0000,0.0000,-150.0000
C02427=20.000,45.800,100.600,0.0000,0.0000,-150.0000
C02428=15.000,45.800,100.600,0.0000,0.0000,-150.0000
C02429=10.000,45.800,100.600,0.0000,0.0000,-150.0000
C02430=5.000,45.800,100.600,0.0000,0.0000,-150.0000
C02431=0.000,45.800,100.600,0.0000,0.0000,-150.0000
C02432=-5.000,45.800,100.600,0.0000,0.0000,-150.0000
C02433=-10.000,45.800,100.600,0.0000,0.0000,-150.0000
C02434=-15.000,45.800,100.600,0.0000,0.0000,-150.0000
C02435=-20.000,45.800,100.600,0.0000,0.0000,-150.0000
C02436=-25.000,45.800,100.600,0.0000,0.0000,-150.0000
C02437=-30.000,45.800,100.600,0.0000,0.0000,-150.0000
C02438=-35.000,45.800,100.600,0.0000,0.0000,-150.0000
C02439=-40.000,45.800,100.600,0.0000,0.0000,-150.0000
C02440=-45.000,45.800,100.600,0.0000,0.0000,-150.0000
C02441=-50.000,45.800,100.600,0.0000,0.0000,-150.0000
C02442=-55.000,45.800,100.600,0.0000,0.0000,-150.0000
C02443=-60.000,45.800,100.600,0.0000,0.0000,-150.0000
C02444=-65.000,45.800,100.600,0.0000,0.0000,-150.0000
C02445=-70.000,45.800,100.600,0.0000,0.0000,-150.0000
C02446=-75.000,45.800,100.600,0.0000,0.0000,-150.0000
C02447=-76.950,43.850,100.600,0.0000,0.0000,-150.0000
C02448=-75.000,41.900,100.600,0.0000,0.0000,-150.0000
C02449=-70.195,41.900,100.600,0.0000,0.0000,-150.0000
C02450=-65.390,41.900,100.600,0.0000,0.0000,-150.0000
C02451=-60.585,41.900,100.600,0.0000,0.0000,-150.0000
C02452=-55.780,41.900,100.600,0.0000,0.0000,-150.0000
C02453=-50.975,41.900,100.600,0.0000,0.0000,-150.0000
C02454=-46.170,41.900,100.600,0.0000,0.0000,-150.0000
C02455=-41.365,41.900,100.600,0.0000,0.0000,-150.0000
C02456=-36.560,41.900,100.600,0.0000,0.0000,-150.0000
C02457=-31.755,41.900,100.600,0.0000,0.0000,-150.0000
C02458=-26.950,41.900,100.600,0.0000,0.0000,-150.0000
C02459=-26.950,36.900,100.600,0.0000,0.0000,-150.0000
C02460=-26.950,31.900,100.600,0.0000,0.0000,-150.0000
C02461=-26.950,26.900,100.600,0.0000,0.0000,-150.0000
C02462=-26.950,21.900,100.600,0.0000,0.0000,-150.0000
C02463=-26.950,16.900,100.600,0.0000,0.0000,-150.0000
C02464=-26.950,11.900,100.600,0.0000,0.0000,-150.0000
C02465=-26.950,6.900,100.600,0.0000,0.0000,-150.0000
C02466=-26.950,1.900,100.600,0.0000,0.0000,-150.0000
C02467=-26.950,-3.100,100.600,0.0000,0.0000,-150.0000
C02468=-26.950,-8.100,100.600,0.0000,0.0000,-150.0000
C02469=-26.950,-13.100,100.600,0.0000,0.0000,-150.0000
C02470=-26.950,-18.100,100.600,0.0000,0.0000,-150.0000
C02471=-26.950,-23.100,100.600,0.0000,0.0000,-150.0000
C02472=-26.950,-28.100,100.600,0.0000,0.0000,-150.0000
C02473=-26.950,-33.100,100.600,0.0000,0.0000,-150.0000
C02474=-26.950,-38.100,100.600,0.0000,0.0000,-150.0000
C02475=-26.950,-43.100,100.600,0.0000,0.0000,-150.0000
C02476=-26.950,-48.100,100.600,0.0000,0.0000,-150.0000
C02477=-26.950,-53.100,100.600,0.0000,0.0000,-150.0000
C02478=-26.950,-58.100,100.600,0.0000,0.0000,-150.0000
C02479=-26.950,-63.100,100.600,0.0000,0.0000,-150.0000
C02480=-26.950,-68.100,100.600,0.0000,0.0000,-150.0000
C02481=-31.755,-68.100,100.600,0.0000,0.0000,-150.0000
C02482=-36.560,-68.100,100.600,0.0000,0.0000,-150.0000
C02483=-41.365,-68.100,100.600,0.0000,0.0000,-150.0000
C02484=-46.170,-68.100,100.600,0.0000,0.0000,-150.0000
C02485=-50.975,-68.100,100.600,0.0000,0.0000,-150.0000
C02486=-55.780,-68.100,100.600,0.0000,0.0000,-150.0000
C02487=-60.585,-68.100,100.600,0.0000,0.0000,-150.0000
C02488=-65.390,-68.100,100.600,0.0000,0.0000,-150.0000
C02489=-70.195,-68.100,100.600,0.0000,0.0000,-150.0000
C02490=-75.000,-68.100,100.600,0.0000,0.0000,-150.0000
C02491=-75.000,-68.100,102.300,0.0000,0.0000,-150.0000
C02492=-70.195,-68.100,102.300,0.0000,0.0000,-150.0000
C02493=-65.390,-68.100,102.300,0.0000,0.0000,-150.0000
C02494=-60.585,-68.100,102.300,0.0000,0.0000,-150.0000
C02495=-55.780,-68.100,102.300,0.0000,0.0000,-150.0000
C02496=-50.975,-68.100,102.300,0.0000,0.0000,-150.0000
C02497=-46.170,-68.100,102.300,0.0000,0.0000,-150.0000
C02498=-41.365,-68.100,102.300,0.0000,0.0000,-150.0000
C02499=-36.560,-68.100,102.300,0.0000,0.0000,-150.0000
C02500=-31.755,-68.100,102.300,0.0000,0.0000,-150.0000
C02501=-26.950,-68.100,102.300,0.0000,0.0000,-150.0000
C02502=-26.950,-63.100,102.300,0.0000,0.0000,-150.0000
C02503=-26.950,-58.100,102.300,0.0000,0.0000,-150.0000
C02504=-26.950,-53.100,102.300,0.0000,0.0000,-150.0000
C02505=-26.950,-48.100,102.300,0.0000,0.0000,-150.0000
C02506=-26.950,-43.100,102.300,0.0000,0.0000,-150.0000
C02507=-26.950,-38.100,102.300,0.0000,0.0000,-150.0000
C02508=-26.950,-33.100,102.300,0.0000,0.0000,-150.0000
C02509=-26.950,-28.100,102.300,0.0000,0.0000,-150.0000
C02510=-26.950,-23.100,102.300,0.0000,0.0000,-150.0000
C02511=-26.950,-18.100,102.300,0.0000,0.0000,-150.0000
C02512=-26.950,-13.100,102.300,0.0000,0.0000,-150.0000
C02513=-26.950,-8.100,102.300,0.0000,0.0000,-150.0000
C02514=-26.950,-3.100,102.300,0.0000,0.0000,-150.0000
C02515=-26.950,1.900,102.300,0.0000,0.0000,-150.0000
C02516=-26.950,6.900,102.300,0.0000,0.0000,-150.0000
C02517=-26.950,11.900,102.300,0.0000,0.0000,-150.0000
C02518=-26.950,16.900,102.300,0.0000,0.0000,-150.0000
C02519=-26.950,21.900,102.300,0.0000,0.0000,-150.0000
C02520=-26.950,26.900,102.300,0.0000,0.0000,-150.0000
C02521=-26.950,31.900,102.300,0.0000,0.0000,-150.0000
C02522=-26.950,36.900,102.300,0.0000,0.0000,-150.0000
C02523=-26.950,41.900,102.300,0.0000,0.0000,-150.0000
C02524=-31.733,41.900,102.300,0.0000,0.0000,-150.0000
C02525=-36.517,41.900,102.300,0.0000,0.0000,-150.0000
C02526=-41.300,41.900,102.300,0.0000,0.0000,-150.0000
C02527=-46.083,41.900,102.300,0.0000,0.0000,-150.0000
C02528=-50.867,41.900,102.300,0.0000,0.0000,-150.0000
C02529=-55.650,41.900,102.300,0.0000,0.0000,-150.0000
C02530=-60.433,41.900,102.300,0.0000,0.0000,-150.0000
C02531=-65.217,41.900,102.300,0.0000,0.0000,-150.0000
C02532=-70.000,41.900,102.300,0.0000,0.0000,-150.0000
C02533=-75.000,41.900,102.300,0.0000,0.0000,-150.0000
C02534=-76.950,43.850,102.300,0.0000,0.0000,-150.0000
C02535=-75.000,45.800,102.300,0.0000,0.0000,-150.0000
C02536=-70.000,45.800,102.300,0.0000,0.0000,-150.0000
C02537=-65.000,45.800,102.300,0.0000,0.0000,-150.0000
C02538=-60.000,45.800,102.300,0.0000,0.0000,-150.0000
C02539=-55.000,45.800,102.300,0.0000,0.0000,-150.0000
C02540=-50.000,45.800,102.300,0.0000,0.0000,-150.0000
C02541=-45.000,45.800,102.300,0.0000,0.0000,-150.0000
C02542=-40.000,45.800,102.300,0.0000,0.0000,-150.0000
C02543=-35.000,45.800,102.300,0.0000,0.0000,-150.0000
C02544=-30.000,45.800,102.300,0.0000,0.0000,-150.0000
C02545=-25.000,45.800,102.300,0.0000,0.0000,-150.0000
C02546=-20.000,45.800,102.300,0.0000,0.0000,-150.0000
C02547=-15.000,45.800,102.300,0.0000,0.0000,-150.0000
C02548=-10.000,45.800,102.300,0.0000,0.0000,-150.0000
C02549=-5.000,45.800,102.300,0.0000,0.0000,-150.0000
C02550=0.000,45.800,102.300,0.0000,0.0000,-150.0000
C02551=5.000,45.800,102.300,0.0000,0.0000,-150.0000
C02552=10.000,45.800,102.300,0.0000,0.0000,-150.0000
C02553=15.000,45.800,102.300,0.0000,0.0000,-150.0000
C02554=20.000,45.800,102.300,0.0000,0.0000,-150.0000
C02555=25.000,45.800,102.300,0.0000,0.0000,-150.0000
C02556=26.950,43.850,102.300,0.0000,0.0000,-150.0000
C02557=25.000,41.900,102.300,0.0000,0.0000,-150.0000
C02558=20.195,41.900,102.300,0.0000,0.0000,-150.0000
C02559=15.390,41.900,102.300,0.0000,0.0000,-150.0000
C02560=10.585,41.900,102.300,0.0000,0.0000,-150.0000
C02561=5.780,41.900,102.300,0.0000,0.0000,-150.0000
C02562=0.975,41.900,102.300,0.0000,0.0000,-150.0000
C02563=-3.830,41.900,102.300,0.0000,0.0000,-150.0000
C02564=-8.635,41.900,102.300,0.0000,0.0000,-150.0000
C02565=-13.440,41.900,102.300,0.0000,0.0000,-150.0000
C02566=-18.245,41.900,102.300,0.0000,0.0000,-150.0000
C02567=-23.050,41.900,102.300,0.0000,0.0000,-150.0000
C02568=-23.050,36.900,102.300,0.0000,0.0000,-150.0000
C02569=-23.050,31.900,102.300,0.0000,0.0000,-150.0000
C02570=-23.050,26.900,102.300,0.0000,0.0000,-150.0000
C02571=-23.050,21.900,102.300,0.0000,0.0000,-150.0000
C02572=-23.050,16.900,102.300,0.0000,0.0000,-150.0000
C02573=-23.050,11.900,102.300,0.0000,0.0000,-150.0000
C02574=-23.050,6.900,102.300,0.0000,0.0000,-150.0000
C02575=-23.050,1.900,102.300,0.0000,0.0000,-150.0000
C02576=-23.050,-3.100,102.300,0.0000,0.0000,-150.0000
C02577=-23.050,-8.100,102.300,0.0000,0.0000,-150.0000
C02578=-23.050,-13.100,102.300,0.0000,0.0000,-150.0000
C02579=-23.050,-18.100,102.300,0.0000,0.0000,-150.0000
C02580=-23.050,-23.100,102.300,0.0000,0.0000,-150.0000
C02581=-23.050,-28.100,102.300,0.0000,0.0000,-150.0000
C02582=-23.050,-33.100,102.300,0.0000,0.0000,-150.0000
C02583=-23.050,-38.100,102.300,0.0000,0.0000,-150.0000
C02584=-23.050,-43.100,102.300,0.0000,0.0000,-150.0000
C02585=-23.050,-48.100,102.300,0.0000,0.0000,-150.0000
C02586=-23.050,-53.100,102.300,0.0000,0.0000,-150.0000
C02587=-23.050,-58.100,102.300,0.0000,0.0000,-150.0000
C02588=-23.050,-63.100,102.300,0.0000,0.0000,-150.0000
C02589=-23.050,-68.100,102.300,0.0000,0.0000,-150.0000
C02590=-18.267,-68.100,102.300,0.0000,0.0000,-150.0000
C02591=-13.483,-68.100,102.300,0.0000,0.0000,-150.0000
C02592=-8.700,-68.100,102.300,0.0000,0.0000,-150.0000
C02593=-3.917,-68.100,102.300,0.0000,0.0000,-150.0000
C02594=0.867,-68.100,102.300,0.0000,0.0000,-150.0000
C02595=5.650,-68.100,102.300,0.0000,0.0000,-150.0000
C02596=10.433,-68.100,102.300,0.0000,0.0000,-150.0000
C02597=15.217,-68.100,102.300,0.0000,0.0000,-150.0000
C02598=20.000,-68.100,102.300,0.0000,0.0000,-150.0000
C02599=25.000,-68.100,102.300,0.0000,0.0000,-150.0000
C02600=26.950,-70.050,102.300,0.0000,0.0000,-150.0000
C02601=25.000,-72.000,102.300,0.0000,0.0000,-150.0000
C02602=20.000,-72.000,102.300,0.0000,0.0000,-150.0000
C02603=15.000,-72.000,102.300,0.0000,0.0000,-150.0000
C02604=10.000,-72.000,102.300,0.0000,0.0000,-150.0000
C02605=5.000,-72.000,102.300,0.0000,0.0000,-150.0000
C02606=0.000,-72.000,102.300,0.0000,0.0000,-150.0000
C02607=-5.000,-72.000,102.300,0.0000,0.0000,-150.0000
C02608=-10.000,-72.000,102.300,0.0000,0.0000,-150.0000
C02609=-15.000,-72.000,102.300,0.0000,0.0000,-150.0000
C02610=-20.000,-72.000,102.300,0.0000,0.0000,-150.0000
C02611=-25.000,-72.000,102.300,0.0000,0.0000,-150.0000
C02612=-30.000,-72.000,102.300,0.0000,0.0000,-150.0000
C02613=-35.000,-72.000,102.300,0.0000,0.0000,-150.0000
C02614=-40.000,-72.000,102.300,0.0000,0.0000,-150.0000
C02615=-45.000,-72.000,102.300,0.0000,0.0000,-150.0000
C02616=-50.000,-72.000,102.300,0.0000,0.0000,-150.0000
C02617=-55.000,-72.000,102.300,0.0000,0.0000,-150.0000
C02618=-60.000,-72.000,102.300,0.0000,0.0000,-150.0000
C02619=-65.000,-72.000,102.300,0.0000,0.0000,-150.0000
C02620=-70.000,-72.000,102.300,0.0000,0.0000,-150.0000
C02621=-75.000,-72.000,102.300,0.0000,0.0000,-150.0000
C02622=-75.000,-72.000,200.000,0.0000,0.0000,-150.0000
C02623=-107.000,-40.000,200.000,0.0000,0.0000,-150.0000
//INST
///DATE 2026/11/26 13:56
///ATTR SC,RW,RJ
////FRAME USER 1
///GROUP1 RB1
NOP
MOVJ C00000 VJ=0.78
MOVJ C00001 VJ=0.78
MOVL C00002 V=11.0 ACC=20 DEC=20
*LAG1
MACRO1 MJ#(0) ARGF1
ARCON
MOVL C00003 V=7.0 ACC=20 DEC=20
MOVL C00004 V=7.0 ACC=20 DEC=20
MOVL C00005 V=7.0 ACC=20 DEC=20
MOVL C00006 V=7.0 ACC=20 DEC=20
MOVL C00007 V=7.0 ACC=20 DEC=20
MOVL C00008 V=7.0 ACC=20 DEC=20
MOVL C00009 V=7.0 ACC=20 DEC=20
MOVL C00010 V=7.0 ACC=20 DEC=20
MOVL C00011 V=7.0 ACC=20 DEC=20
MOVL C00012 V=7.0 ACC=20 DEC=20
MOVL C00013 V=7.0 ACC=20 DEC=20
MOVL C00014 V=7.0 ACC=20 DEC=20
MOVL C00015 V=7.0 ACC=20 DEC=20
MOVL C00016 V=7.0 ACC=20 DEC=20
MOVL C00017 V=7.0 ACC=20 DEC=20
MOVL C00018 V=7.0 ACC=20 DEC=20
MOVL C00019 V=7.0 ACC=20 DEC=20
MOVL C00020 V=7.0 ACC=20 DEC=20
MOVL C00021 V=7.0 ACC=20 DEC=20
MOVC C00022 V=12.0 ACC=20 DEC=20
MOVC C00023 V=12.0 ACC=20 DEC=20
MOVC C00024 V=12.0 ACC=20 DEC=20
MOVL C00025 V=7.0 ACC=20 DEC=20
MOVL C00026 V=7.0 ACC=20 DEC=20
MOVL C00027 V=7.0 ACC=20 DEC=20
MOVL C00028 V=7.0 ACC=20 DEC=20
MOVL C00029 V=7.0 ACC=20 DEC=20
MOVL C00030 V=7.0 ACC=20 DEC=20
MOVL C00031 V=7.0 ACC=20 DEC=20
MOVL C00032 V=7.0 ACC=20 DEC=20
MOVL C00033 V=7.0 ACC=20 DEC=20
MOVL C00034 V=7.0 PL=1
MOVL C00035 V=7.0 ACC=20 DEC=20
MOVL C00036 V=7.0 ACC=20 DEC=20
MOVL C00037 V=7.0 ACC=20 DEC=20
MOVL C00038 V=7.0 ACC=20 DEC=20
MOVL C00039 V=7.0 ACC=20 DEC=20
MOVL C00040 V=7.0 ACC=20 DEC=20
MOVL C00041 V=7.0 ACC=20 DEC=20
MOVL C00042 V=7.0 ACC=20 DEC=20
MOVL C00043 V=7.0 ACC=20 DEC=20
MOVL C00044 V=7.0 ACC=20 DEC=20
MOVL C00045 V=7.0 ACC=20 DEC=20
MOVL C00046 V=7.0 ACC=20 DEC=20
MOVL C00047 V=7.0 ACC=20 DEC=20
MOVL C00048 V=7.0 ACC=20 DEC=20
MOVL C00049 V=7.0 ACC=20 DEC=20
MOVL C00050 V=7.0 ACC=20 DEC=20
MOVL C00051 V=7.0 ACC=20 DEC=20
MOVL C00052 V=7.0 ACC=20 DEC=20
MOVL C00053 V=7.0 ACC=20 DEC=20
MOVL C00054 V=7.0 ACC=20 DEC=20
MOVL C00055 V=7.0 ACC=20 DEC=20
MOVL C00056 V=7.0 PL=1
MOVL C00057 V=7.0 ACC=20 DEC=20
MOVL C00058 V=7.0 ACC=20 DEC=20
MOVL C00059 V=7.0 ACC=20 DEC=20
MOVL C00060 V=7.0 ACC=20 DEC=20
MOVL C00061 V=7.0 ACC=20 DEC=20
MOVL C00062 V=7.0 ACC=20 DEC=20
MOVL C00063 V=7.0 ACC=20 DEC=20
MOVL C00064 V=7.0 ACC=20 DEC=20
MOVL C00065 V=7.0 ACC=20 DEC=20
MOVC C00066 V=12.0 ACC=20 DEC=20
MOVC C00067 V=12.0 ACC=20 DEC=20
MOVC C00068 V=12.0 ACC=20 DEC=20
MOVL C00069 V=7.0 ACC=20 DEC=20
MOVL C00070 V=7.0 ACC=20 DEC=20
MOVL C00071 V=7.0 ACC=20 DEC=20
MOVL C00072 V=7.0 ACC=20 DEC=20
MOVL C00073 V=7.0 ACC=20 DEC=20
MOVL C00074 V=7.0 ACC=20 DEC=20
MOVL C00075 V=7.0 ACC=20 DEC=20
MOVL C00076 V=7.0 ACC=20 DEC=20
MOVL C00077 V=7.0 ACC=20 DEC=20
MOVL C00078 V=7.0 ACC=20 DEC=20
MOVL C00079 V=7.0 ACC=20 DEC=20
MOVL C00080 V=7.0 ACC=20 DEC=20
MOVL C00081 V=7.0 ACC=20 DEC=20
MOVL C00082 V=7.0 ACC=20 DEC=20
MOVL C00083 V=7.0 ACC=20 DEC=20
MOVL C00084 V=7.0 ACC=20 DEC=20
MOVL C00085 V=7.0 ACC=20 DEC=20
MOVL C00086 V=7.0 ACC=20 DEC=20
MOVL C00087 V=7.0 ACC=20 DEC=20
MOVC C00088 V=12.0 ACC=20 DEC=20
MOVC C00089 V=12.0 ACC=20 DEC=20
MOVC C00090 V=12.0 ACC=20 DEC=20
MOVL C00091 V=7.0 ACC=20 DEC=20
MOVL C00092 V=7.0 ACC=20 DEC=20
MOVL C00093 V=7.0 ACC=20 DEC=20
MOVL C00094 V=7.0 ACC=20 DEC=20
MOVL C00095 V=7.0 ACC=20 DEC=20
MOVL C00096 V=7.0 ACC=20 DEC=20
MOVL C00097 V=7.0 ACC=20 DEC=20
MOVL C00098 V=7.0 ACC=20 DEC=20
MOVL C00099 V=7.0 ACC=20 DEC=20
MOVL C00100 V=7.0 PL=1
MOVL C00101 V=7.0 ACC=20 DEC=20
MOVL C00102 V=7.0 ACC=20 DEC=20
MOVL C00103 V=7.0 ACC=20 DEC=20
MOVL C00104 V=7.0 ACC=20 DEC=20
MOVL C00105 V=7.0 ACC=20 DEC=20
MOVL C00106 V=7.0 ACC=20 DEC=20
MOVL C00107 V=7.0 ACC=20 DEC=20
MOVL C00108 V=7.0 ACC=20 DEC=20
MOVL C00109 V=7.0 ACC=20 DEC=20
MOVL C00110 V=7.0 ACC=20 DEC=20
MOVL C00111 V=7.0 ACC=20 DEC=20
MOVL C00112 V=7.0 ACC=20 DEC=20
MOVL C00113 V=7.0 ACC=20 DEC=20
MOVL C00114 V=7.0 ACC=20 DEC=20
MOVL C00115 V=7.0 ACC=20 DEC=20
MOVL C00116 V=7.0 ACC=20 DEC=20
MOVL C00117 V=7.0 ACC=20 DEC=20
MOVL C00118 V=7.0 ACC=20 DEC=20
MOVL C00119 V=7.0 ACC=20 DEC=20
MOVL C00120 V=7.0 ACC=20 DEC=20
MOVL C00121 V=7.0 ACC=20 DEC=20
MOVL C00122 V=7.0 PL=1
MOVL C00123 V=7.0 ACC=20 DEC=20
MOVL C00124 V=7.0 ACC=20 DEC=20
MOVL C00125 V=7.0 ACC=20 DEC=20
MOVL C00126 V=7.0 ACC=20 DEC=20
MOVL C00127 V=7.0 ACC=20 DEC=20
MOVL C00128 V=7.0 ACC=20 DEC=20
MOVL C00129 V=7.0 ACC=20 DEC=20
MOVL C00130 V=7.0 ACC=20 DEC=20
MOVL C00131 V=7.0 ACC=20 DEC=20
MOVL C00132 V=7.0 ACC=20 DEC=20
ARCOF
TIMER T=30
MOVL C00133 V=11.0 ACC=20 DEC=20
*LAG2
MACRO1 MJ#(0) ARGF2
ARCON
MOVL C00134 V=7.0 ACC=20 DEC=20
MOVL C00135 V=7.0 ACC=20 DEC=20
MOVL C00136 V=7.0 ACC=20 DEC=20
MOVL C00137 V=7.0 ACC=20 DEC=20
MOVL C00138 V=7.0 ACC=20 DEC=20
MOVL C00139 V=7.0 ACC=20 DEC=20
MOVL C00140 V=7.0 ACC=20 DEC=20
MOVL C00141 V=7.0 ACC=20 DEC=20
MOVL C00142 V=7.0 ACC=20 DEC=20
MOVL C00143 V=7.0 PL=1
MOVL C00144 V=7.0 ACC=20 DEC=20
MOVL C00145 V=7.0 ACC=20 DEC=20
MOVL C00146 V=7.0 ACC=20 DEC=20
MOVL C00147 V=7.0 ACC=20 DEC=20
MOVL C00148 V=7.0 ACC=20 DEC=20
MOVL C00149 V=7.0 ACC=20 DEC=20
MOVL C00150 V=7.0 ACC=20 DEC=20
MOVL C00151 V=7.0 ACC=20 DEC=20
MOVL C00152 V=7.0 ACC=20 DEC=20
MOVL C00153 V=7.0 ACC=20 DEC=20
MOVL C00154 V=7.0 ACC=20 DEC=20
MOVL C00155 V=7.0 ACC=20 DEC=20
MOVL C00156 V=7.0 ACC=20 DEC=20
MOVL C00157 V=7.0 ACC=20 DEC=20
MOVL C00158 V=7.0 ACC=20 DEC=20
MOVL C00159 V=7.0 ACC=20 DEC=20
MOVL C00160 V=7.0 ACC=20 DEC=20
MOVL C00161 V=7.0 ACC=20 DEC=20
MOVL C00162 V=7.0 ACC=20 DEC=20
MOVL C00163 V=7.0 ACC=20 DEC=20
MOVL C00164 V=7.0 ACC=20 DEC=20
MOVL C00165 V=7.0 PL=1
MOVL C00166 V=7.0 ACC=20 DEC=20
MOVL C00167 V=7.0 ACC=20 DEC=20
MOVL C00168 V=7.0 ACC=20 DEC=20
MOVL C00169 V=7.0 ACC=20 DEC=20
MOVL C00170 V=7.0 ACC=20 DEC=20
MOVL C00171 V=7.0 ACC=20 DEC=20
MOVL C00172 V=7.0 ACC=20 DEC=20
MOVL C00173 V=7.0 ACC=20 DEC=20
MOVL C00174 V=7.0 ACC=20 DEC=20
MOVC C00175 V=12.0 ACC=20 DEC=20
MOVC C00176 V=12.0 ACC=20 DEC=20
MOVC C00177 V=12.0 ACC=20 DEC=20
MOVL C00178 V=7.0 ACC=20 DEC=20
MOVL C00179 V=7.0 ACC=20 DEC=20
MOVL C00180 V=7.0 ACC=20 DEC=20
MOVL C00181 V=7.0 ACC=20 DEC=20
MOVL C00182 V=7.0 ACC=20 DEC=20
MOVL C00183 V=7.0 ACC=20 DEC=20
MOVL C00184 V=7.0 ACC=20 DEC=20
MOVL C00185 V=7.0 ACC=20 DEC=20
MOVL C00186 V=7.0 ACC=20 DEC=20
MOVL C00187 V=7.0 ACC=20 DEC=20
MOVL C00188 V=7.0 ACC=20 DEC=20
MOVL C00189 V=7.0 ACC=20 DEC=20
MOVL C00190 V=7.0 ACC=20 DEC=20
MOVL C00191 V=7.0 ACC=20 DEC=20
MOVL C00192 V=7.0 ACC=20 DEC=20
MOVL C00193 V=7.0 ACC=20 DEC=20
MOVL C00194 V=7.0 ACC=20 DEC=20
MOVL C00195 V=7.0 ACC=20 DEC=20
MOVL C00196 V=7.0 ACC=20 DEC=20
MOVC C00197 V=12.0 ACC=20 DEC=20
MOVC C00198 V=12.0 ACC=20 DEC=20
MOVC C00199 V=12.0 ACC=20 DEC=20
MOVL C00200 V=7.0 ACC=20 DEC=20
MOVL C00201 V=7.0 ACC=20 DEC=20
MOVL C00202 V=7.0 ACC=20 DEC=20
MOVL C00203 V=7.0 ACC=20 DEC=20
MOVL C00204 V=7.0 ACC=20 DEC=20
MOVL C00205 V=7.0 ACC=20 DEC=20
MOVL C00206 V=7.0 ACC=20 DEC=20
MOVL C00207 V=7.0 ACC=20 DEC=20
MOVL C00208 V=7.0 ACC=20 DEC=20
MOVL C00209 V=7.0 PL=1
MOVL C00210 V=7.0 ACC=20 DEC=20
MOVL C00211 V=7.0 ACC=20 DEC=20
MOVL C00212 V=7.0 ACC=20 DEC=20
MOVL C00213 V=7.0 ACC=20 DEC=20
MOVL C00214 V=7.0 ACC=20 DEC=20
MOVL C00215 V=7.0 ACC=20 DEC=20
MOVL C00216 V=7.0 ACC=20 DEC=20
MOVL C00217 V=7.0 ACC=20 DEC=20
MOVL C00218 V=7.0 ACC=20 DEC=20
MOVL C00219 V=7.0 ACC=20 DEC=20
MOVL C00220 V=7.0 ACC=20 DEC=20
MOVL C00221 V=7.0 ACC=20 DEC=20
MOVL C00222 V=7.0 ACC=20 DEC=20
MOVL C00223 V=7.0 ACC=20 DEC=20
MOVL C00224 V=7.0 ACC=20 DEC=20
MOVL C00225 V=7.0 ACC=20 DEC=20
MOVL C00226 V=7.0 ACC=20 DEC=20
MOVL C00227 V=7.0 ACC=20 DEC=20
MOVL C00228 V=7.0 ACC=20 DEC=20
MOVL C00229 V=7.0 ACC=20 DEC=20
MOVL C00230 V=7.0 ACC=20 DEC=20
MOVL C00231 V=7.0 PL=1
MOVL C00232 V=7.0 ACC=20 DEC=20
MOVL C00233 V=7.0 ACC=20 DEC=20
MOVL C00234 V=7.0 ACC=20 DEC=20
MOVL C00235 V=7.0 ACC=20 DEC=20
MOVL C00236 V=7.0 ACC=20 DEC=20
MOVL C00237 V=7.0 ACC=20 DEC=20
MOVL C00238 V=7.0 ACC=20 DEC=20
MOVL C00239 V=7.0 ACC=20 DEC=20
MOVL C00240 V=7.0 ACC=20 DEC=20
MOVC C00241 V=12.0 ACC=20 DEC=20
MOVC C00242 V=12.0 ACC=20 DEC=20
MOVC C00243 V=12.0 ACC=20 DEC=20
MOVL C00244 V=7.0 ACC=20 DEC=20
MOVL C00245 V=7.0 ACC=20 DEC=20
MOVL C00246 V=7.0 ACC=20 DEC=20
MOVL C00247 V=7.0 ACC=20 DEC=20
MOVL C00248 V=7.0 ACC=20 DEC=20
MOVL C00249 V=7.0 ACC=20 DEC=20
MOVL C00250 V=7.0 ACC=20 DEC=20
MOVL C00251 V=7.0 ACC=20 DEC=20
MOVL C00252 V=7.0 ACC=20 DEC=20
MOVL C00253 V=7.0 ACC=20 DEC=20
MOVL C00254 V=7.0 ACC=20 DEC=20
MOVL C00255 V=7.0 ACC=20 DEC=20
MOVL C00256 V=7.0 ACC=20 DEC=20
MOVL C00257 V=7.0 ACC=20 DEC=20
MOVL C00258 V=7.0 ACC=20 DEC=20
MOVL C00259 V=7.0 ACC=20 DEC=20
MOVL C00260 V=7.0 ACC=20 DEC=20
MOVL C00261 V=7.0 ACC=20 DEC=20
MOVL C00262 V=7.0 ACC=20 DEC=20
MOVL C00263 V=7.0 ACC=20 DEC=20
ARCOF
TIMER T=30
MOVL C00264 V=11.0 ACC=20 DEC=20
*LAG3
MACRO1 MJ#(0) ARGF2
ARCON
MOVL C00265 V=7.0 ACC=20 DEC=20
MOVL C00266 V=7.0 ACC=20 DEC=20
MOVL C00267 V=7.0 ACC=20 DEC=20
MOVL C00268 V=7.0 ACC=20 DEC=20
MOVL C00269 V=7.0 ACC=20 DEC=20
MOVL C00270 V=7.0 ACC=20 DEC=20
MOVL C00271 V=7.0 ACC=20 DEC=20
MOVL C00272 V=7.0 ACC=20 DEC=20
MOVL C00273 V=7.0 ACC=20 DEC=20
MOVL C00274 V=7.0 ACC=20 DEC=20
MOVL C00275 V=7.0 ACC=20 DEC=20
MOVL C00276 V=7.0 ACC=20 DEC=20
MOVL C00277 V=7.0 ACC=20 DEC=20
MOVL C00278 V=7.0 ACC=20 DEC=20
MOVL C00279 V=7.0 ACC=20 DEC=20
MOVL C00280 V=7.0 ACC=20 DEC=20
MOVL C00281 V=7.0 ACC=20 DEC=20
MOVL C00282 V=7.0 ACC=20 DEC=20
MOVL C00283 V=7.0 ACC=20 DEC=20
MOVC C00284 V=12.0 ACC=20 DEC=20
MOVC C00285 V=12.0 ACC=20 DEC=20
MOVC C00286 V=12.0 ACC=20 DEC=20
MOVL C00287 V=7.0 ACC=20 DEC=20
MOVL C00288 V=7.0 ACC=20 DEC=20
MOVL C00289 V=7.0 ACC=20 DEC=20
MOVL C00290 V=7.0 ACC=20 DEC=20
MOVL C00291 V=7.0 ACC=20 DEC=20
MOVL C00292 V=7.0 ACC=20 DEC=20
MOVL C00293 V=7.0 ACC=20 DEC=20
MOVL C00294 V=7.0 ACC=20 DEC=20
MOVL C00295 V=7.0 ACC=20 DEC=20
MOVL C00296 V=7.0 PL=1
MOVL C00297 V=7.0 ACC=20 DEC=20
MOVL C00298 V=7.0 ACC=20 DEC=20
MOVL C00299 V=7.0 ACC=20 DEC=20
MOVL C00300 V=7.0 ACC=20 DEC=20
MOVL C00301 V=7.0 ACC=20 DEC=20
MOVL C00302 V=7.0 ACC=20 DEC=20
MOVL C00303 V=7.0 ACC=20 DEC=20
MOVL C00304 V=7.0 ACC=20 DEC=20
MOVL C00305 V=7.0 ACC=20 DEC=20
MOVL C00306 V=7.0 ACC=20 DEC=20
MOVL C00307 V=7.0 ACC=20 DEC=20
MOVL C00308 V=7.0 ACC=20 DEC=20
MOVL C00309 V=7.0 ACC=20 DEC=20
MOVL C00310 V=7.0 ACC=20 DEC=20
MOVL C00311 V=7.0 ACC=20 DEC=20
MOVL C00312 V=7.0 ACC=20 DEC=20
MOVL C00313 V=7.0 ACC=20 DEC=20
MOVL C00314 V=7.0 ACC=20 DEC=20
MOVL C00315 V=7.0 ACC=20 DEC=20
MOVL C00316 V=7.0 ACC=20 DEC=20
MOVL C00317 V=7.0 ACC=20 DEC=20
MOVL C00318 V=7.0 PL=1
MOVL C00319 V=7.0 ACC=20 DEC=20
MOVL C00320 V=7.0 ACC=20 DEC=20
MOVL C00321 V=7.0 ACC=20 DEC=20
MOVL C00322 V=7.0 ACC=20 DEC=20
MOVL C00323 V=7.0 ACC=20 DEC=20
MOVL C00324 V=7.0 ACC=20 DEC=20
MOVL C00325 V=7.0 ACC=20 DEC=20
MOVL C00326 V=7.0 ACC=20 DEC=20
MOVL C00327 V=7.0 ACC=20 DEC=20
MOVC C00328 V=12.0 ACC=20 DEC=20
MOVC C00329 V=12.0 ACC=20 DEC=20
MOVC C00330 V=12.0 ACC=20 DEC=20
MOVL C00331 V=7.0 ACC=20 DEC=20
MOVL C00332 V=7.0 ACC=20 DEC=20
MOVL C00333 V=7.0 ACC=20 DEC=20
MOVL C00334 V=7.0 ACC=20 DEC=20
MOVL C00335 V=7.0 ACC=20 DEC=20
MOVL C00336 V=7.0 ACC=20 DEC=20
MOVL C00337 V=7.0 ACC=20 DEC=20
MOVL C00338 V=7.0 ACC=20 DEC=20
MOVL C00339 V=7.0 ACC=20 DEC=20
MOVL C00340 V=7.0 ACC=20 DEC=20
MOVL C00341 V=7.0 ACC=20 DEC=20
MOVL C00342 V=7.0 ACC=20 DEC=20
MOVL C00343 V=7.0 ACC=20 DEC=20
MOVL C00344 V=7.0 ACC=20 DEC=20
MOVL C00345 V=7.0 ACC=20 DEC=20
MOVL C00346 V=7.0 ACC=20 DEC=20
MOVL C00347 V=7.0 ACC=20 DEC=20
MOVL C00348 V=7.0 ACC=20 DEC=20
MOVL C00349 V=7.0 ACC=20 DEC=20
MOVC C00350 V=12.0 ACC=20 DEC=20
MOVC C00351 V=12.0 ACC=20 DEC=20
MOVC C00352 V=12.0 ACC=20 DEC=20
MOVL C00353 V=7.0 ACC=20 DEC=20
MOVL C00354 V=7.0 ACC=20 DEC=20
MOVL C00355 V=7.0 ACC=20 DEC=20
MOVL C00356 V=7.0 ACC=20 DEC=20
MOVL C00357 V=7.0 ACC=20 DEC=20
MOVL C00358 V=7.0 ACC=20 DEC=20
MOVL C00359 V=7.0 ACC=20 DEC=20
MOVL C00360 V=7.0 ACC=20 DEC=20
MOVL C00361 V=7.0 ACC=20 DEC=20
MOVL C00362 V=7.0 PL=1
MOVL C00363 V=7.0 ACC=20 DEC=20
MOVL C00364 V=7.0 ACC=20 DEC=20
MOVL C00365 V=7.0 ACC=20 DEC=20
MOVL C00366 V=7.0 ACC=20 DEC=20
MOVL C00367 V=7.0 ACC=20 DEC=20
MOVL C00368 V=7.0 ACC=20 DEC=20
MOVL C00369 V=7.0 ACC=20 DEC=20
MOVL C00370 V=7.0 ACC=20 DEC=20
MOVL C00371 V=7.0 ACC=20 DEC=20
MOVL C00372 V=7.0 ACC=20 DEC=20
MOVL C00373 V=7.0 ACC=20 DEC=20
MOVL C00374 V=7.0 ACC=20 DEC=20
MOVL C00375 V=7.0 ACC=20 DEC=20
MOVL C00376 V=7.0 ACC=20 DEC=20
MOVL C00377 V=7.0 ACC=20 DEC=20
MOVL C00378 V=7.0 ACC=20 DEC=20
MOVL C00379 V=7.0 ACC=20 DEC=20
MOVL C00380 V=7.0 ACC=20 DEC=20
MOVL C00381 V=7.0 ACC=20 DEC=20
MOVL C00382 V=7.0 ACC=20 DEC=20
MOVL C00383 V=7.0 ACC=20 DEC=20
MOVL C00384 V=7.0 PL=1
MOVL C00385 V=7.0 ACC=20 DEC=20
MOVL C00386 V=7.0 ACC=20 DEC=20
MOVL C00387 V=7.0 ACC=20 DEC=20
MOVL C00388 V=7.0 ACC=20 DEC=20
MOVL C00389 V=7.0 ACC=20 DEC=20
MOVL C00390 V=7.0 ACC=20 DEC=20
MOVL C00391 V=7.0 ACC=20 DEC=20
MOVL C00392 V=7.0 ACC=20 DEC=20
MOVL C00393 V=7.0 ACC=20 DEC=20
MOVL C00394 V=7.0 ACC=20 DEC=20
ARCOF
TIMER T=30
MOVL C00395 V=11.0 ACC=20 DEC=20
*LAG4
MACRO1 MJ#(0) ARGF2
ARCON
MOVL C00396 V=7.0 ACC=20 DEC=20
MOVL C00397 V=7.0 ACC=20 DEC=20
MOVL C00398 V=7.0 ACC=20 DEC=20
MOVL C00399 V=7.0 ACC=20 DEC=20
MOVL C00400 V=7.0 ACC=20 DEC=20
MOVL C00401 V=7.0 ACC=20 DEC=20
MOVL C00402 V=7.0 ACC=20 DEC=20
MOVL C00403 V=7.0 ACC=20 DEC=20
MOVL C00404 V=7.0 ACC=20 DEC=20
MOVL C00405 V=7.0 PL=1
MOVL C00406 V=7.0 ACC=20 DEC=20
MOVL C00407 V=7.0 ACC=20 DEC=20
MOVL C00408 V=7.0 ACC=20 DEC=20
MOVL C00409 V=7.0 ACC=20 DEC=20
MOVL C00410 V=7.0 ACC=20 DEC=20
MOVL C00411 V=7.0 ACC=20 DEC=20
MOVL C00412 V=7.0 ACC=20 DEC=20
MOVL C00413 V=7.0 ACC=20 DEC=20
MOVL C00414 V=7.0 ACC=20 DEC=20
MOVL C00415 V=7.0 ACC=20 DEC=20
MOVL C00416 V=7.0 ACC=20 DEC=20
MOVL C00417 V=7.0 ACC=20 DEC=20
MOVL C00418 V=7.0 ACC=20 DEC=20
MOVL C00419 V=7.0 ACC=20 DEC=20
MOVL C00420 V=7.0 ACC=20 DEC=20
MOVL C00421 V=7.0 ACC=20 DEC=20
MOVL C00422 V=7.0 ACC=20 DEC=20
MOVL C00423 V=7.0 ACC=20 DEC=20
MOVL C00424 V=7.0 ACC=20 DEC=20
MOVL C00425 V=7.0 ACC=20 DEC=20
MOVL C00426 V=7.0 ACC=20 DEC=20
MOVL C00427 V=7.0 PL=1
MOVL C00428 V=7.0 ACC=20 DEC=20
MOVL C00429 V=7.0 ACC=20 DEC=20
MOVL C00430 V=7.0 ACC=20 DEC=20
MOVL C00431 V=7.0 ACC=20 DEC=20
MOVL C00432 V=7.0 ACC=20 DEC=20
MOVL C00433 V=7.0 ACC=20 DEC=20
MOVL C00434 V=7.0 ACC=20 DEC=20
MOVL C00435 V=7.0 ACC=20 DEC=20
MOVL C00436 V=7.0 ACC=20 DEC=20
MOVC C00437 V=12.0 ACC=20 DEC=20
MOVC C00438 V=12.0 ACC=20 DEC=20
MOVC C00439 V=12.0 ACC=20 DEC=20
MOVL C00440 V=7.0 ACC=20 DEC=20
MOVL C00441 V=7.0 ACC=20 DEC=20
MOVL C00442 V=7.0 ACC=20 DEC=20
MOVL C00443 V=7.0 ACC=20 DEC=20
MOVL C00444 V=7.0 ACC=20 DEC=20
MOVL C00445 V=7.0 ACC=20 DEC=20
MOVL C00446 V=7.0 ACC=20 DEC=20
MOVL C00447 V=7.0 ACC=20 DEC=20
MOVL C00448 V=7.0 ACC=20 DEC=20
MOVL C00449 V=7.0 ACC=20 DEC=20
MOVL C00450 V=7.0 ACC=20 DEC=20
MOVL C00451 V=7.0 ACC=20 DEC=20
MOVL C00452 V=7.0 ACC=20 DEC=20
MOVL C00453 V=7.0 ACC=20 DEC=20
MOVL C00454 V=7.0 ACC=20 DEC=20
MOVL C00455 V=7.0 ACC=20 DEC=20
MOVL C00456 V=7.0 ACC=20 DEC=20
MOVL C00457 V=7.0 ACC=20 DEC=20
MOVL C00458 V=7.0 ACC=20 DEC=20
MOVC C00459 V=12.0 ACC=20 DEC=20
MOVC C00460 V=12.0 ACC=20 DEC=20
MOVC C00461 V=12.0 ACC=20 DEC=20
MOVL C00462 V=7.0 ACC=20 DEC=20
MOVL C00463 V=7.0 ACC=20 DEC=20
MOVL C00464 V=7.0 ACC=20 DEC=20
MOVL C00465 V=7.0 ACC=20 DEC=20
MOVL C00466 V=7.0 ACC=20 DEC=20
MOVL C00467 V=7.0 ACC=20 DEC=20
MOVL C00468 V=7.0 ACC=20 DEC=20
MOVL C00469 V=7.0 ACC=20 DEC=20
MOVL C00470 V=7.0 ACC=20 DEC=20
MOVL C00471 V=7.0 PL=1
MOVL C00472 V=7.0 ACC=20 DEC=20
MOVL C00473 V=7.0 ACC=20 DEC=20
MOVL C00474 V=7.0 ACC=20 DEC=20
MOVL C00475 V=7.0 ACC=20 DEC=20
MOVL C00476 V=7.0 ACC=20 DEC=20
MOVL C00477 V=7.0 ACC=20 DEC=20
MOVL C00478 V=7.0 ACC=20 DEC=20
MOVL C00479 V=7.0 ACC=20 DEC=20
MOVL C00480 V=7.0 ACC=20 DEC=20
MOVL C00481 V=7.0 ACC=20 DEC=20
MOVL C00482 V=7.0 ACC=20 DEC=20
MOVL C00483 V=7.0 ACC=20 DEC=20
MOVL C00484 V=7.0 ACC=20 DEC=20
MOVL C00485 V=7.0 ACC=20 DEC=20
MOVL C00486 V=7.0 ACC=20 DEC=20
MOVL C00487 V=7.0 ACC=20 DEC=20
MOVL C00488 V=7.0 ACC=20 DEC=20
MOVL C00489 V=7.0 ACC=20 DEC=20
MOVL C00490 V=7.0 ACC=20 DEC=20
MOVL C00491 V=7.0 ACC=20 DEC=20
MOVL C00492 V=7.0 ACC=20 DEC=20
MOVL C00493 V=7.0 PL=1
MOVL C00494 V=7.0 ACC=20 DEC=20
MOVL C00495 V=7.0 ACC=20 DEC=20
MOVL C00496 V=7.0 ACC=20 DEC=20
MOVL C00497 V=7.0 ACC=20 DEC=20
MOVL C00498 V=7.0 ACC=20 DEC=20
MOVL C00499 V=7.0 ACC=20 DEC=20
MOVL C00500 V=7.0 ACC=20 DEC=20
MOVL C00501 V=7.0 ACC=20 DEC=20
MOVL C00502 V=7.0 ACC=20 DEC=20
MOVC C00503 V=12.0 ACC=20 DEC=20
MOVC C00504 V=12.0 ACC=20 DEC=20
MOVC C00505 V=12.0 ACC=20 DEC=20
MOVL C00506 V=7.0 ACC=20 DEC=20
MOVL C00507 V=7.0 ACC=20 DEC=20
MOVL C00508 V=7.0 ACC=20 DEC=20
MOVL C00509 V=7.0 ACC=20 DEC=20
MOVL C00510 V=7.0 ACC=20 DEC=20
MOVL C00511 V=7.0 ACC=20 DEC=20
MOVL C00512 V=7.0 ACC=20 DEC=20
MOVL C00513 V=7.0 ACC=20 DEC=20
MOVL C00514 V=7.0 ACC=20 DEC=20
MOVL C00515 V=7.0 ACC=20 DEC=20
MOVL C00516 V=7.0 ACC=20 DEC=20
MOVL C00517 V=7.0 ACC=20 DEC=20
MOVL C00518 V=7.0 ACC=20 DEC=20
MOVL C00519 V=7.0 ACC=20 DEC=20
MOVL C00520 V=7.0 ACC=20 DEC=20
MOVL C00521 V=7.0 ACC=20 DEC=20
MOVL C00522 V=7.0 ACC=20 DEC=20
MOVL C00523 V=7.0 ACC=20 DEC=20
MOVL C00524 V=7.0 ACC=20 DEC=20
MOVL C00525 V=7.0 ACC=20 DEC=20
ARCOF
TIMER T=30
MOVL C00526 V=11.0 ACC=20 DEC=20
*LAG5
MACRO1 MJ#(0) ARGF2
ARCON
MOVL C00527 V=7.0 ACC=20 DEC=20
MOVL C00528 V=7.0 ACC=20 DEC=20
MOVL C00529 V=7.0 ACC=20 DEC=20
MOVL C00530 V=7.0 ACC=20 DEC=20
MOVL C00531 V=7.0 ACC=20 DEC=20
MOVL C00532 V=7.0 ACC=20 DEC=20
MOVL C00533 V=7.0 ACC=20 DEC=20
MOVL C00534 V=7.0 ACC=20 DEC=20
MOVL C00535 V=7.0 ACC=20 DEC=20
MOVL C00536 V=7.0 ACC=20 DEC=20
MOVL C00537 V=7.0 ACC=20 DEC=20
MOVL C00538 V=7.0 ACC=20 DEC=20
MOVL C00539 V=7.0 ACC=20 DEC=20
MOVL C00540 V=7.0 ACC=20 DEC=20
MOVL C00541 V=7.0 ACC=20 DEC=20
MOVL C00542 V=7.0 ACC=20 DEC=20
MOVL C00543 V=7.0 ACC=20 DEC=20
MOVL C00544 V=7.0 ACC=20 DEC=20
MOVL C00545 V=7.0 ACC=20 DEC=20
MOVC C00546 V=12.0 ACC=20 DEC=20
MOVC C00547 V=12.0 ACC=20 DEC=20
MOVC C00548 V=12.0 ACC=20 DEC=20
MOVL C00549 V=7.0 ACC=20 DEC=20
MOVL C00550 V=7.0 ACC=20 DEC=20
MOVL C00551 V=7.0 ACC=20 DEC=20
MOVL C00552 V=7.0 ACC=20 DEC=20
MOVL C00553 V=7.0 ACC=20 DEC=20
MOVL C00554 V=7.0 ACC=20 DEC=20
MOVL C00555 V=7.0 ACC=20 DEC=20
MOVL C00556 V=7.0 ACC=20 DEC=20
MOVL C00557 V=7.0 ACC=20 DEC=20
MOVL C00558 V=7.0 PL=1
MOVL C00559 V=7.0 ACC=20 DEC=20
MOVL C00560 V=7.0 ACC=20 DEC=20
MOVL C00561 V=7.0 ACC=20 DEC=20
MOVL C00562 V=7.0 ACC=20 DEC=20
MOVL C00563 V=7.0 ACC=20 DEC=20
MOVL C00564 V=7.0 ACC=20 DEC=20
MOVL C00565 V=7.0 ACC=20 DEC=20
MOVL C00566 V=7.0 ACC=20 DEC=20
MOVL C00567 V=7.0 ACC=20 DEC=20
MOVL C00568 V=7.0 ACC=20 DEC=20
MOVL C00569 V=7.0 ACC=20 DEC=20
MOVL C00570 V=7.0 ACC=20 DEC=20
MOVL C00571 V=7.0 ACC=20 DEC=20
MOVL C00572 V=7.0 ACC=20 DEC=20
MOVL C00573 V=7.0 ACC=20 DEC=20
MOVL C00574 V=7.0 ACC=20 DEC=20
MOVL C00575 V=7.0 ACC=20 DEC=20
MOVL C00576 V=7.0 ACC=20 DEC=20
MOVL C00577 V=7.0 ACC=20 DEC=20
MOVL C00578 V=7.0 ACC=20 DEC=20
MOVL C00579 V=7.0 ACC=20 DEC=20
MOVL C00580 V=7.0 PL=1
MOVL C00581 V=7.0 ACC=20 DEC=20
MOVL C00582 V=7.0 ACC=20 DEC=20
MOVL C00583 V=7.0 ACC=20 DEC=20
MOVL C00584 V=7.0 ACC=20 DEC=20
MOVL C00585 V=7.0 ACC=20 DEC=20
MOVL C00586 V=7.0 ACC=20 DEC=20
MOVL C00587 V=7.0 ACC=20 DEC=20
MOVL C00588 V=7.0 ACC=20 DEC=20
MOVL C00589 V=7.0 ACC=20 DEC=20
MOVC C00590 V=12.0 ACC=20 DEC=20
MOVC C00591 V=12.0 ACC=20 DEC=20
MOVC C00592 V=12.0 ACC=20 DEC=20
MOVL C00593 V=7.0 ACC=20 DEC=20
MOVL C00594 V=7.0 ACC=20 DEC=20
MOVL C00595 V=7.0 ACC=20 DEC=20
MOVL C00596 V=7.0 ACC=20 DEC=20
MOVL C00597 V=7.0 ACC=20 DEC=20
MOVL C00598 V=7.0 ACC=20 DEC=20
MOVL C00599 V=7.0 ACC=20 DEC=20
MOVL C00600 V=7.0 ACC=20 DEC=20
MOVL C00601 V=7.0 ACC=20 DEC=20
MOVL C00602 V=7.0 ACC=20 DEC=20
MOVL C00603 V=7.0 ACC=20 DEC=20
MOVL C00604 V=7.0 ACC=20 DEC=20
MOVL C00605 V=7.0 ACC=20 DEC=20
MOVL C00606 V=7.0 ACC=20 DEC=20
MOVL C00607 V=7.0 ACC=20 DEC=20
MOVL C00608 V=7.0 ACC=20 DEC=20
MOVL C00609 V=7.0 ACC=20 DEC=20
MOVL C00610 V=7.0 ACC=20 DEC=20
MOVL C00611 V=7.0 ACC=20 DEC=20
MOVC C00612 V=12.0 ACC=20 DEC=20
MOVC C00613 V=12.0 ACC=20 DEC=20
MOVC C00614 V=12.0 ACC=20 DEC=20
MOVL C00615 V=7.0 ACC=20 DEC=20
MOVL C00616 V=7.0 ACC=20 DEC=20
MOVL C00617 V=7.0 ACC=20 DEC=20
MOVL C00618 V=7.0 ACC=20 DEC=20
MOVL C00619 V=7.0 ACC=20 DEC=20
MOVL C00620 V=7.0 ACC=20 DEC=20
MOVL C00621 V=7.0 ACC=20 DEC=20
MOVL C00622 V=7.0 ACC=20 DEC=20
MOVL C00623 V=7.0 ACC=20 DEC=20
MOVL C00624 V=7.0 PL=1
MOVL C00625 V=7.0 ACC=20 DEC=20
MOVL C00626 V=7.0 ACC=20 DEC=20
MOVL C00627 V=7.0 ACC=20 DEC=20
MOVL C00628 V=7.0 ACC=20 DEC=20
MOVL C00629 V=7.0 ACC=20 DEC=20
MOVL C00630 V=7.0 ACC=20 DEC=20
MOVL C00631 V=7.0 ACC=20 DEC=20
MOVL C00632 V=7.0 ACC=20 DEC=20
MOVL C00633 V=7.0 ACC=20 DEC=20
MOVL C00634 V=7.0 ACC=20 DEC=20
MOVL C00635 V=7.0 ACC=20 DEC=20
MOVL C00636 V=7.0 ACC=20 DEC=20
MOVL C00637 V=7.0 ACC=20 DEC=20
MOVL C00638 V=7.0 ACC=20 DEC=20
MOVL C00639 V=7.0 ACC=20 DEC=20
MOVL C00640 V=7.0 ACC=20 DEC=20
MOVL C00641 V=7.0 ACC=20 DEC=20
MOVL C00642 V=7.0 ACC=20 DEC=20
MOVL C00643 V=7.0 ACC=20 DEC=20
MOVL C00644 V=7.0 ACC=20 DEC=20
MOVL C00645 V=7.0 ACC=20 DEC=20
MOVL C00646 V=7.0 PL=1
MOVL C00647 V=7.0 ACC=20 DEC=20
MOVL C00648 V=7.0 ACC=20 DEC=20
MOVL C00649 V=7.0 ACC=20 DEC=20
MOVL C00650 V=7.0 ACC=20 DEC=20
MOVL C00651 V=7.0 ACC=20 DEC=20
MOVL C00652 V=7.0 ACC=20 DEC=20
MOVL C00653 V=7.0 ACC=20 DEC=20
MOVL C00654 V=7.0 ACC=20 DEC=20
MOVL C00655 V=7.0 ACC=20 DEC=20
MOVL C00656 V=7.0 ACC=20 DEC=20
ARCOF
TIMER T=30
MOVL C00657 V=11.0 ACC=20 DEC=20
*LAG6
MACRO1 MJ#(0) ARGF2
ARCON
MOVL C00658 V=7.0 ACC=20 DEC=20
MOVL C00659 V=7.0 ACC=20 DEC=20
MOVL C00660 V=7.0 ACC=20 DEC=20
MOVL C00661 V=7.0 ACC=20 DEC=20
MOVL C00662 V=7.0 ACC=20 DEC=20
MOVL C00663 V=7.0 ACC=20 DEC=20
MOVL C00664 V=7.0 ACC=20 DEC=20
MOVL C00665 V=7.0 ACC=20 DEC=20
MOVL C00666 V=7.0 ACC=20 DEC=20
MOVL C00667 V=7.0 PL=1
MOVL C00668 V=7.0 ACC=20 DEC=20
MOVL C00669 V=7.0 ACC=20 DEC=20
MOVL C00670 V=7.0 ACC=20 DEC=20
MOVL C00671 V=7.0 ACC=20 DEC=20
MOVL C00672 V=7.0 ACC=20 DEC=20
MOVL C00673 V=7.0 ACC=20 DEC=20
MOVL C00674 V=7.0 ACC=20 DEC=20
MOVL C00675 V=7.0 ACC=20 DEC=20
MOVL C00676 V=7.0 ACC=20 DEC=20
MOVL C00677 V=7.0 ACC=20 DEC=20
MOVL C00678 V=7.0 ACC=20 DEC=20
MOVL C00679 V=7.0 ACC=20 DEC=20
MOVL C00680 V=7.0 ACC=20 DEC=20
MOVL C00681 V=7.0 ACC=20 DEC=20
MOVL C00682 V=7.0 ACC=20 DEC=20
MOVL C00683 V=7.0 ACC=20 DEC=20
MOVL C00684 V=7.0 ACC=20 DEC=20
MOVL C00685 V=7.0 ACC=20 DEC=20
MOVL C00686 V=7.0 ACC=20 DEC=20
MOVL C00687 V=7.0 ACC=20 DEC=20
MOVL C00688 V=7.0 ACC=20 DEC=20
MOVL C00689 V=7.0 PL=1
MOVL C00690 V=7.0 ACC=20 DEC=20
MOVL C00691 V=7.0 ACC=20 DEC=20
MOVL C00692 V=7.0 ACC=20 DEC=20
MOVL C00693 V=7.0 ACC=20 DEC=20
MOVL C00694 V=7.0 ACC=20 DEC=20
MOVL C00695 V=7.0 ACC=20 DEC=20
MOVL C00696 V=7.0 ACC=20 DEC=20
MOVL C00697 V=7.0 ACC=20 DEC=20
MOVL C00698 V=7.0 ACC=20 DEC=20
MOVC C00699 V=12.0 ACC=20 DEC=20
MOVC C00700 V=12.0 ACC=20 DEC=20
MOVC C00701 V=12.0 ACC=20 DEC=20
MOVL C00702 V=7.0 ACC=20 DEC=20
MOVL C00703 V=7.0 ACC=20 DEC=20
MOVL C00704 V=7.0 ACC=20 DEC=20
MOVL C00705 V=7.0 ACC=20 DEC=20
MOVL C00706 V=7.0 ACC=20 DEC=20
MOVL C00707 V=7.0 ACC=20 DEC=20
MOVL C00708 V=7.0 ACC=20 DEC=20
MOVL C00709 V=7.0 ACC=20 DEC=20
MOVL C00710 V=7.0 ACC=20 DEC=20
MOVL C00711 V=7.0 ACC=20 DEC=20
MOVL C00712 V=7.0 ACC=20 DEC=20
MOVL C00713 V=7.0 ACC=20 DEC=20
MOVL C00714 V=7.0 ACC=20 DEC=20
MOVL C00715 V=7.0 ACC=20 DEC=20
MOVL C00716 V=7.0 ACC=20 DEC=20
MOVL C00717 V=7.0 ACC=20 DEC=20
MOVL C00718 V=7.0 ACC=20 DEC=20
MOVL C00719 V=7.0 ACC=20 DEC=20
MOVL C00720 V=7.0 ACC=20 DEC=20
MOVC C00721 V=12.0 ACC=20 DEC=20
MOVC C00722 V=12.0 ACC=20 DEC=20
MOVC C00723 V=12.0 ACC=20 DEC=20
MOVL C00724 V=7.0 ACC=20 DEC=20
MOVL C00725 V=7.0 ACC=20 DEC=20
MOVL C00726 V=7.0 ACC=20 DEC=20
MOVL C00727 V=7.0 ACC=20 DEC=20
MOVL C00728 V=7.0 ACC=20 DEC=20
MOVL C00729 V=7.0 ACC=20 DEC=20
MOVL C00730 V=7.0 ACC=20 DEC=20
MOVL C00731 V=7.0 ACC=20 DEC=20
MOVL C00732 V=7.0 ACC=20 DEC=20
MOVL C00733 V=7.0 PL=1
MOVL C00734 V=7.0 ACC=20 DEC=20
MOVL C00735 V=7.0 ACC=20 DEC=20
MOVL C00736 V=7.0 ACC=20 DEC=20
MOVL C00737 V=7.0 ACC=20 DEC=20
MOVL C00738 V=7.0 ACC=20 DEC=20
MOVL C00739 V=7.0 ACC=20 DEC=20
MOVL C00740 V=7.0 ACC=20 DEC=20
MOVL C00741 V=7.0 ACC=20 DEC=20
MOVL C00742 V=7.0 ACC=20 DEC=20
MOVL C00743 V=7.0 ACC=20 DEC=20
MOVL C00744 V=7.0 ACC=20 DEC=20
MOVL C00745 V=7.0 ACC=20 DEC=20
MOVL C00746 V=7.0 ACC=20 DEC=20
MOVL C00747 V=7.0 ACC=20 DEC=20
MOVL C00748 V=7.0 ACC=20 DEC=20
MOVL C00749 V=7.0 ACC=20 DEC=20
MOVL C00750 V=7.0 ACC=20 DEC=20
MOVL C00751 V=7.0 ACC=20 DEC=20
MOVL C00752 V=7.0 ACC=20 DEC=20
MOVL C00753 V=7.0 ACC=20 DEC=20
MOVL C00754 V=7.0 ACC=20 DEC=20
MOVL C00755 V=7.0 PL=1
MOVL C00756 V=7.0 ACC=20 DEC=20
MOVL C00757 V=7.0 ACC=20 DEC=20
MOVL C00758 V=7.0 ACC=20 DEC=20
MOVL C00759 V=7.0 ACC=20 DEC=20
MOVL C00760 V=7.0 ACC=20 DEC=20
MOVL C00761 V=7.0 ACC=20 DEC=20
MOVL C00762 V=7.0 ACC=20 DEC=20
MOVL C00763 V=7.0 ACC=20 DEC=20
MOVL C00764 V=7.0 ACC=20 DEC=20
MOVC C00765 V=12.0 ACC=20 DEC=20
MOVC C00766 V=12.0 ACC=20 DEC=20
MOVC C00767 V=12.0 ACC=20 DEC=20
MOVL C00768 V=7.0 ACC=20 DEC=20
MOVL C00769 V=7.0 ACC=20 DEC=20
MOVL C00770 V=7.0 ACC=20 DEC=20
MOVL C00771 V=7.0 ACC=20 DEC=20
MOVL C00772 V=7.0 ACC=20 DEC=20
MOVL C00773 V=7.0 ACC=20 DEC=20
MOVL C00774 V=7.0 ACC=20 DEC=20
MOVL C00775 V=7.0 ACC=20 DEC=20
MOVL C00776 V=7.0 ACC=20 DEC=20
MOVL C00777 V=7.0 ACC=20 DEC=20
MOVL C00778 V=7.0 ACC=20 DEC=20
MOVL C00779 V=7.0 ACC=20 DEC=20
MOVL C00780 V=7.0 ACC=20 DEC=20
MOVL C00781 V=7.0 ACC=20 DEC=20
MOVL C00782 V=7.0 ACC=20 DEC=20
MOVL C00783 V=7.0 ACC=20 DEC=20
MOVL C00784 V=7.0 ACC=20 DEC=20
MOVL C00785 V=7.0 ACC=20 DEC=20
MOVL C00786 V=7.0 ACC=20 DEC=20
MOVL C00787 V=7.0 ACC=20 DEC=20
ARCOF
TIMER T=30
MOVL C00788 V=11.0 ACC=20 DEC=20
*LAG7
MACRO1 MJ#(0) ARGF2
ARCON
MOVL C00789 V=7.0 ACC=20 DEC=20
MOVL C00790 V=7.0 ACC=20 DEC=20
MOVL C00791 V=7.0 ACC=20 DEC=20
MOVL C00792 V=7.0 ACC=20 DEC=20
MOVL C00793 V=7.0 ACC=20 DEC=20
MOVL C00794 V=7.0 ACC=20 DEC=20
MOVL C00795 V=7.0 ACC=20 DEC=20
MOVL C00796 V=7.0 ACC=20 DEC=20
MOVL C00797 V=7.0 ACC=20 DEC=20
MOVL C00798 V=7.0 ACC=20 DEC=20
MOVL C00799 V=7.0 ACC=20 DEC=20
MOVL C00800 V=7.0 ACC=20 DEC=20
MOVL C00801 V=7.0 ACC=20 DEC=20
MOVL C00802 V=7.0 ACC=20 DEC=20
MOVL C00803 V=7.0 ACC=20 DEC=20
MOVL C00804 V=7.0 ACC=20 DEC=20
MOVL C00805 V=7.0 ACC=20 DEC=20
MOVL C00806 V=7.0 ACC=20 DEC=20
MOVL C00807 V=7.0 ACC=20 DEC=20
MOVC C00808 V=12.0 ACC=20 DEC=20
MOVC C00809 V=12.0 ACC=20 DEC=20
MOVC C00810 V=12.0 ACC=20 DEC=20
MOVL C00811 V=7.0 ACC=20 DEC=20
MOVL C00812 V=7.0 ACC=20 DEC=20
MOVL C00813 V=7.0 ACC=20 DEC=20
MOVL C00814 V=7.0 ACC=20 DEC=20
MOVL C00815 V=7.0 ACC=20 DEC=20
MOVL C00816 V=7.0 ACC=20 DEC=20
MOVL C00817 V=7.0 ACC=20 DEC=20
MOVL C00818 V=7.0 ACC=20 DEC=20
MOVL C00819 V=7.0 ACC=20 DEC=20
MOVL C00820 V=7.0 PL=1
MOVL C00821 V=7.0 ACC=20 DEC=20
MOVL C00822 V=7.0 ACC=20 DEC=20
MOVL C00823 V=7.0 ACC=20 DEC=20
MOVL C00824 V=7.0 ACC=20 DEC=20
MOVL C00825 V=7.0 ACC=20 DEC=20
MOVL C00826 V=7.0 ACC=20 DEC=20
MOVL C00827 V=7.0 ACC=20 DEC=20
MOVL C00828 V=7.0 ACC=20 DEC=20
MOVL C00829 V=7.0 ACC=20 DEC=20
MOVL C00830 V=7.0 ACC=20 DEC=20
MOVL C00831 V=7.0 ACC=20 DEC=20
MOVL C00832 V=7.0 ACC=20 DEC=20
MOVL C00833 V=7.0 ACC=20 DEC=20
MOVL C00834 V=7.0 ACC=20 DEC=20
MOVL C00835 V=7.0 ACC=20 DEC=20
MOVL C00836 V=7.0 ACC=20 DEC=20
MOVL C00837 V=7.0 ACC=20 DEC=20
MOVL C00838 V=7.0 ACC=20 DEC=20
MOVL C00839 V=7.0 ACC=20 DEC=20
MOVL C00840 V=7.0 ACC=20 DEC=20
MOVL C00841 V=7.0 ACC=20 DEC=20
MOVL C00842 V=7.0 PL=1
MOVL C00843 V=7.0 ACC=20 DEC=20
MOVL C00844 V=7.0 ACC=20 DEC=20
MOVL C00845 V=7.0 ACC=20 DEC=20
MOVL C00846 V=7.0 ACC=20 DEC=20
MOVL C00847 V=7.0 ACC=20 DEC=20
MOVL C00848 V=7.0 ACC=20 DEC=20
MOVL C00849 V=7.0 ACC=20 DEC=20
MOVL C00850 V=7.0 ACC=20 DEC=20
MOVL C00851 V=7.0 ACC=20 DEC=20
MOVC C00852 V=12.0 ACC=20 DEC=20
MOVC C00853 V=12.0 ACC=20 DEC=20
MOVC C00854 V=12.0 ACC=20 DEC=20
MOVL C00855 V=7.0 ACC=20 DEC=20
MOVL C00856 V=7.0 ACC=20 DEC=20
MOVL C00857 V=7.0 ACC=20 DEC=20
MOVL C00858 V=7.0 ACC=20 DEC=20
MOVL C00859 V=7.0 ACC=20 DEC=20
MOVL C00860 V=7.0 ACC=20 DEC=20
MOVL C00861 V=7.0 ACC=20 DEC=20
MOVL C00862 V=7.0 ACC=20 DEC=20
MOVL C00863 V=7.0 ACC=20 DEC=20
MOVL C00864 V=7.0 ACC=20 DEC=20
MOVL C00865 V=7.0 ACC=20 DEC=20
MOVL C00866 V=7.0 ACC=20 DEC=20
MOVL C00867 V=7.0 ACC=20 DEC=20
MOVL C00868 V=7.0 ACC=20 DEC=20
MOVL C00869 V=7.0 ACC=20 DEC=20
MOVL C00870 V=7.0 ACC=20 DEC=20
MOVL C00871 V=7.0 ACC=20 DEC=20
MOVL C00872 V=7.0 ACC=20 DEC=20
MOVL C00873 V=7.0 ACC=20 DEC=20
MOVC C00874 V=12.0 ACC=20 DEC=20
MOVC C00875 V=12.0 ACC=20 DEC=20
MOVC C00876 V=12.0 ACC=20 DEC=20
MOVL C00877 V=7.0 ACC=20 DEC=20
MOVL C00878 V=7.0 ACC=20 DEC=20
MOVL C00879 V=7.0 ACC=20 DEC=20
MOVL C00880 V=7.0 ACC=20 DEC=20
MOVL C00881 V=7.0 ACC=20 DEC=20
MOVL C00882 V=7.0 ACC=20 DEC=20
MOVL C00883 V=7.0 ACC=20 DEC=20
MOVL C00884 V=7.0 ACC=20 DEC=20
MOVL C00885 V=7.0 ACC=20 DEC=20
MOVL C00886 V=7.0 PL=1
MOVL C00887 V=7.0 ACC=20 DEC=20
MOVL C00888 V=7.0 ACC=20 DEC=20
MOVL C00889 V=7.0 ACC=20 DEC=20
MOVL C00890 V=7.0 ACC=20 DEC=20
MOVL C00891 V=7.0 ACC=20 DEC=20
MOVL C00892 V=7.0 ACC=20 DEC=20
MOVL C00893 V=7.0 ACC=20 DEC=20
MOVL C00894 V=7.0 ACC=20 DEC=20
MOVL C00895 V=7.0 ACC=20 DEC=20
MOVL C00896 V=7.0 ACC=20 DEC=20
MOVL C00897 V=7.0 ACC=20 DEC=20
MOVL C00898 V=7.0 ACC=20 DEC=20
MOVL C00899 V=7.0 ACC=20 DEC=20
MOVL C00900 V=7.0 ACC=20 DEC=20
MOVL C00901 V=7.0 ACC=20 DEC=20
MOVL C00902 V=7.0 ACC=20 DEC=20
MOVL C00903 V=7.0 ACC=20 DEC=20
MOVL C00904 V=7.0 ACC=20 DEC=20
MOVL C00905 V=7.0 ACC=20 DEC=20
MOVL C00906 V=7.0 ACC=20 DEC=20
MOVL C00907 V=7.0 ACC=20 DEC=20
MOVL C00908 V=7.0 PL=1
MOVL C00909 V=7.0 ACC=20 DEC=20
MOVL C00910 V=7.0 ACC=20 DEC=20
MOVL C00911 V=7.0 ACC=20 DEC=20
MOVL C00912 V=7.0 ACC=20 DEC=20
MOVL C00913 V=7.0 ACC=20 DEC=20
MOVL C00914 V=7.0 ACC=20 DEC=20
MOVL C00915 V=7.0 ACC=20 DEC=20
MOVL C00916 V=7.0 ACC=20 DEC=20
MOVL C00917 V=7.0 ACC=20 DEC=20
MOVL C00918 V=7.0 ACC=20 DEC=20
ARCOF
TIMER T=30
MOVL C00919 V=11.0 ACC=20 DEC=20
*LAG8
MACRO1 MJ#(0) ARGF2
ARCON
MOVL C00920 V=7.0 ACC=20 DEC=20
MOVL C00921 V=7.0 ACC=20 DEC=20
MOVL C00922 V=7.0 ACC=20 DEC=20
MOVL C00923 V=7.0 ACC=20 DEC=20
MOVL C00924 V=7.0 ACC=20 DEC=20
MOVL C00925 V=7.0 ACC=20 DEC=20
MOVL C00926 V=7.0 ACC=20 DEC=20
MOVL C00927 V=7.0 ACC=20 DEC=20
MOVL C00928 V=7.0 ACC=20 DEC=20
MOVL C00929 V=7.0 PL=1
MOVL C00930 V=7.0 ACC=20 DEC=20
MOVL C00931 V=7.0 ACC=20 DEC=20
MOVL C00932 V=7.0 ACC=20 DEC=20
MOVL C00933 V=7.0 ACC=20 DEC=20
MOVL C00934 V=7.0 ACC=20 DEC=20
MOVL C00935 V=7.0 ACC=20 DEC=20
MOVL C00936 V=7.0 ACC=20 DEC=20
MOVL C00937 V=7.0 ACC=20 DEC=20
MOVL C00938 V=7.0 ACC=20 DEC=20
MOVL C00939 V=7.0 ACC=20 DEC=20
MOVL C00940 V=7.0 ACC=20 DEC=20
MOVL C00941 V=7.0 ACC=20 DEC=20
MOVL C00942 V=7.0 ACC=20 DEC=20
MOVL C00943 V=7.0 ACC=20 DEC=20
MOVL C00944 V=7.0 ACC=20 DEC=20
MOVL C00945 V=7.0 ACC=20 DEC=20
MOVL C00946 V=7.0 ACC=20 DEC=20
MOVL C00947 V=7.0 ACC=20 DEC=20
MOVL C00948 V=7.0 ACC=20 DEC=20
MOVL C00949 V=7.0 ACC=20 DEC=20
MOVL C00950 V=7.0 ACC=20 DEC=20
MOVL C00951 V=7.0 PL=1
MOVL C00952 V=7.0 ACC=20 DEC=20
MOVL C00953 V=7.0 ACC=20 DEC=20
MOVL C00954 V=7.0 ACC=20 DEC=20
MOVL C00955 V=7.0 ACC=20 DEC=20
MOVL C00956 V=7.0 ACC=20 DEC=20
MOVL C00957 V=7.0 ACC=20 DEC=20
MOVL C00958 V=7.0 ACC=20 DEC=20
MOVL C00959 V=7.0 ACC=20 DEC=20
MOVL C00960 V=7.0 ACC=20 DEC=20
MOVC C00961 V=12.0 ACC=20 DEC=20
MOVC C00962 V=12.0 ACC=20 DEC=20
MOVC C00963 V=12.0 ACC=20 DEC=20
MOVL C00964 V=7.0 ACC=20 DEC=20
MOVL C00965 V=7.0 ACC=20 DEC=20
MOVL C00966 V=7.0 ACC=20 DEC=20
MOVL C00967 V=7.0 ACC=20 DEC=20
MOVL C00968 V=7.0 ACC=20 DEC=20
MOVL C00969 V=7.0 ACC=20 DEC=20
MOVL C00970 V=7.0 ACC=20 DEC=20
MOVL C00971 V=7.0 ACC=20 DEC=20
MOVL C00972 V=7.0 ACC=20 DEC=20
MOVL C00973 V=7.0 ACC=20 DEC=20
MOVL C00974 V=7.0 ACC=20 DEC=20
MOVL C00975 V=7.0 ACC=20 DEC=20
MOVL C00976 V=7.0 ACC=20 DEC=20
MOVL C00977 V=7.0 ACC=20 DEC=20
MOVL C00978 V=7.0 ACC=20 DEC=20
MOVL C00979 V=7.0 ACC=20 DEC=20
MOVL C00980 V=7.0 ACC=20 DEC=20
MOVL C00981 V=7.0 ACC=20 DEC=20
MOVL C00982 V=7.0 ACC=20 DEC=20
MOVC C00983 V=12.0 ACC=20 DEC=20
MOVC C00984 V=12.0 ACC=20 DEC=20
MOVC C00985 V=12.0 ACC=20 DEC=20
MOVL C00986 V=7.0 ACC=20 DEC=20
MOVL C00987 V=7.0 ACC=20 DEC=20
MOVL C00988 V=7.0 ACC=20 DEC=20
MOVL C00989 V=7.0 ACC=20 DEC=20
MOVL C00990 V=7.0 ACC=20 DEC=20
MOVL C00991 V=7.0 ACC=20 DEC=20
MOVL C00992 V=7.0 ACC=20 DEC=20
MOVL C00993 V=7.0 ACC=20 DEC=20
MOVL C00994 V=7.0 ACC=20 DEC=20
MOVL C00995 V=7.0 PL=1
MOVL C00996 V=7.0 ACC=20 DEC=20
MOVL C00997 V=7.0 ACC=20 DEC=20
MOVL C00998 V=7.0 ACC=20 DEC=20
MOVL C00999 V=7.0 ACC=20 DEC=20
MOVL C01000 V=7.0 ACC=20 DEC=20
MOVL C01001 V=7.0 ACC=20 DEC=20
MOVL C01002 V=7.0 ACC=20 DEC=20
MOVL C01003 V=7.0 ACC=20 DEC=20
MOVL C01004 V=7.0 ACC=20 DEC=20
MOVL C01005 V=7.0 ACC=20 DEC=20
MOVL C01006 V=7.0 ACC=20 DEC=20
MOVL C01007 V=7.0 ACC=20 DEC=20
MOVL C01008 V=7.0 ACC=20 DEC=20
MOVL C01009 V=7.0 ACC=20 DEC=20
MOVL C01010 V=7.0 ACC=20 DEC=20
MOVL C01011 V=7.0 ACC=20 DEC=20
MOVL C01012 V=7.0 ACC=20 DEC=20
MOVL C01013 V=7.0 ACC=20 DEC=20
MOVL C01014 V=7.0 ACC=20 DEC=20
MOVL C01015 V=7.0 ACC=20 DEC=20
MOVL C01016 V=7.0 ACC=20 DEC=20
MOVL C01017 V=7.0 PL=1
MOVL C01018 V=7.0 ACC=20 DEC=20
MOVL C01019 V=7.0 ACC=20 DEC=20
MOVL C01020 V=7.0 ACC=20 DEC=20
MOVL C01021 V=7.0 ACC=20 DEC=20
MOVL C01022 V=7.0 ACC=20 DEC=20
MOVL C01023 V=7.0 ACC=20 DEC=20
MOVL C01024 V=7.0 ACC=20 DEC=20
MOVL C01025 V=7.0 ACC=20 DEC=20
MOVL C01026 V=7.0 ACC=20 DEC=20
MOVC C01027 V=12.0 ACC=20 DEC=20
MOVC C01028 V=12.0 ACC=20 DEC=20
MOVC C01029 V=12.0 ACC=20 DEC=20
MOVL C01030 V=7.0 ACC=20 DEC=20
MOVL C01031 V=7.0 ACC=20 DEC=20
MOVL C01032 V=7.0 ACC=20 DEC=20
MOVL C01033 V=7.0 ACC=20 DEC=20
MOVL C01034 V=7.0 ACC=20 DEC=20
MOVL C01035 V=7.0 ACC=20 DEC=20
MOVL C01036 V=7.0 ACC=20 DEC=20
MOVL C01037 V=7.0 ACC=20 DEC=20
MOVL C01038 V=7.0 ACC=20 DEC=20
MOVL C01039 V=7.0 ACC=20 DEC=20
MOVL C01040 V=7.0 ACC=20 DEC=20
MOVL C01041 V=7.0 ACC=20 DEC=20
MOVL C01042 V=7.0 ACC=20 DEC=20
MOVL C01043 V=7.0 ACC=20 DEC=20
MOVL C01044 V=7.0 ACC=20 DEC=20
MOVL C01045 V=7.0 ACC=20 DEC=20
MOVL C01046 V=7.0 ACC=20 DEC=20
MOVL C01047 V=7.0 ACC=20 DEC=20
MOVL C01048 V=7.0 ACC=20 DEC=20
MOVL C01049 V=7.0 ACC=20 DEC=20
ARCOF
TIMER T=30
MOVL C01050 V=11.0 ACC=20 DEC=20
*LAG9
MACRO1 MJ#(0) ARGF2
ARCON
MOVL C01051 V=7.0 ACC=20 DEC=20
MOVL C01052 V=7.0 ACC=20 DEC=20
MOVL C01053 V=7.0 ACC=20 DEC=20
MOVL C01054 V=7.0 ACC=20 DEC=20
MOVL C01055 V=7.0 ACC=20 DEC=20
MOVL C01056 V=7.0 ACC=20 DEC=20
MOVL C01057 V=7.0 ACC=20 DEC=20
MOVL C01058 V=7.0 ACC=20 DEC=20
MOVL C01059 V=7.0 ACC=20 DEC=20
MOVL C01060 V=7.0 ACC=20 DEC=20
MOVL C01061 V=7.0 ACC=20 DEC=20
MOVL C01062 V=7.0 ACC=20 DEC=20
MOVL C01063 V=7.0 ACC=20 DEC=20
MOVL C01064 V=7.0 ACC=20 DEC=20
MOVL C01065 V=7.0 ACC=20 DEC=20
MOVL C01066 V=7.0 ACC=20 DEC=20
MOVL C01067 V=7.0 ACC=20 DEC=20
MOVL C01068 V=7.0 ACC=20 DEC=20
MOVL C01069 V=7.0 ACC=20 DEC=20
MOVC C01070 V=12.0 ACC=20 DEC=20
MOVC C01071 V=12.0 ACC=20 DEC=20
MOVC C01072 V=12.0 ACC=20 DEC=20
MOVL C01073 V=7.0 ACC=20 DEC=20
MOVL C01074 V=7.0 ACC=20 DEC=20
MOVL C01075 V=7.0 ACC=20 DEC=20
MOVL C01076 V=7.0 ACC=20 DEC=20
MOVL C01077 V=7.0 ACC=20 DEC=20
MOVL C01078 V=7.0 ACC=20 DEC=20
MOVL C01079 V=7.0 ACC=20 DEC=20
MOVL C01080 V=7.0 ACC=20 DEC=20
MOVL C01081 V=7.0 ACC=20 DEC=20
MOVL C01082 V=7.0 PL=1
MOVL C01083 V=7.0 ACC=20 DEC=20
MOVL C01084 V=7.0 ACC=20 DEC=20
MOVL C01085 V=7.0 ACC=20 DEC=20
MOVL C01086 V=7.0 ACC=20 DEC=20
MOVL C01087 V=7.0 ACC=20 DEC=20
MOVL C01088 V=7.0 ACC=20 DEC=20
MOVL C01089 V=7.0 ACC=20 DEC=20
MOVL C01090 V=7.0 ACC=20 DEC=20
MOVL C01091 V=7.0 ACC=20 DEC=20
MOVL C01092 V=7.0 ACC=20 DEC=20
MOVL C01093 V=7.0 ACC=20 DEC=20
MOVL C01094 V=7.0 ACC=20 DEC=20
MOVL C01095 V=7.0 ACC=20 DEC=20
MOVL C01096 V=7.0 ACC=20 DEC=20
MOVL C01097 V=7.0 ACC=20 DEC=20
MOVL C01098 V=7.0 ACC=20 DEC=20
MOVL C01099 V=7.0 ACC=20 DEC=20
MOVL C01100 V=7.0 ACC=20 DEC=20
MOVL C01101 V=7.0 ACC=20 DEC=20
MOVL C01102 V=7.0 ACC=20 DEC=20
MOVL C01103 V=7.0 ACC=20 DEC=20
MOVL C01104 V=7.0 PL=1
MOVL C01105 V=7.0 ACC=20 DEC=20
MOVL C01106 V=7.0 ACC=20 DEC=20
MOVL C01107 V=7.0 ACC=20 DEC=20
MOVL C01108 V=7.0 ACC=20 DEC=20
MOVL C01109 V=7.0 ACC=20 DEC=20
MOVL C01110 V=7.0 ACC=20 DEC=20
MOVL C01111 V=7.0 ACC=20 DEC=20
MOVL C01112 V=7.0 ACC=20 DEC=20
MOVL C01113 V=7.0 ACC=20 DEC=20
MOVC C01114 V=12.0 ACC=20 DEC=20
MOVC C01115 V=12.0 ACC=20 DEC=20
MOVC C01116 V=12.0 ACC=20 DEC=20
MOVL C01117 V=7.0 ACC=20 DEC=20
MOVL C01118 V=7.0 ACC=20 DEC=20
MOVL C01119 V=7.0 ACC=20 DEC=20
MOVL C01120 V=7.0 ACC=20 DEC=20
MOVL C01121 V=7.0 ACC=20 DEC=20
MOVL C01122 V=7.0 ACC=20 DEC=20
MOVL C01123 V=7.0 ACC=20 DEC=20
MOVL C01124 V=7.0 ACC=20 DEC=20
MOVL C01125 V=7.0 ACC=20 DEC=20
MOVL C01126 V=7.0 ACC=20 DEC=20
MOVL C01127 V=7.0 ACC=20 DEC=20
MOVL C01128 V=7.0 ACC=20 DEC=20
MOVL C01129 V=7.0 ACC=20 DEC=20
MOVL C01130 V=7.0 ACC=20 DEC=20
MOVL C01131 V=7.0 ACC=20 DEC=20
MOVL C01132 V=7.0 ACC=20 DEC=20
MOVL C01133 V=7.0 ACC=20 DEC=20
MOVL C01134 V=7.0 ACC=20 DEC=20
MOVL C01135 V=7.0 ACC=20 DEC=20
MOVC C01136 V=12.0 ACC=20 DEC=20
MOVC C01137 V=12.0 ACC=20 DEC=20
MOVC C01138 V=12.0 ACC=20 DEC=20
MOVL C01139 V=7.0 ACC=20 DEC=20
MOVL C01140 V=7.0 ACC=20 DEC=20
MOVL C01141 V=7.0 ACC=20 DEC=20
MOVL C01142 V=7.0 ACC=20 DEC=20
MOVL C01143 V=7.0 ACC=20 DEC=20
MOVL C01144 V=7.0 ACC=20 DEC=20
MOVL C01145 V=7.0 ACC=20 DEC=20
MOVL C01146 V=7.0 ACC=20 DEC=20
MOVL C01147 V=7.0 ACC=20 DEC=20
MOVL C01148 V=7.0 PL=1
MOVL C01149 V=7.0 ACC=20 DEC=20
MOVL C01150 V=7.0 ACC=20 DEC=20
MOVL C01151 V=7.0 ACC=20 DEC=20
MOVL C01152 V=7.0 ACC=20 DEC=20
MOVL C01153 V=7.0 ACC=20 DEC=20
MOVL C01154 V=7.0 ACC=20 DEC=20
MOVL C01155 V=7.0 ACC=20 DEC=20
MOVL C01156 V=7.0 ACC=20 DEC=20
MOVL C01157 V=7.0 ACC=20 DEC=20
MOVL C01158 V=7.0 ACC=20 DEC=20
MOVL C01159 V=7.0 ACC=20 DEC=20
MOVL C01160 V=7.0 ACC=20 DEC=20
MOVL C01161 V=7.0 ACC=20 DEC=20
MOVL C01162 V=7.0 ACC=20 DEC=20
MOVL C01163 V=7.0 ACC=20 DEC=20
MOVL C01164 V=7.0 ACC=20 DEC=20
MOVL C01165 V=7.0 ACC=20 DEC=20
MOVL C01166 V=7.0 ACC=20 DEC=20
MOVL C01167 V=7.0 ACC=20 DEC=20
MOVL C01168 V=7.0 ACC=20 DEC=20
MOVL C01169 V=7.0 ACC=20 DEC=20
MOVL C01170 V=7.0 PL=1
MOVL C01171 V=7.0 ACC=20 DEC=20
MOVL C01172 V=7.0 ACC=20 DEC=20
MOVL C01173 V=7.0 ACC=20 DEC=20
MOVL C01174 V=7.0 ACC=20 DEC=20
MOVL C01175 V=7.0 ACC=20 DEC=20
MOVL C01176 V=7.0 ACC=20 DEC=20
MOVL C01177 V=7.0 ACC=20 DEC=20
MOVL C01178 V=7.0 ACC=20 DEC=20
MOVL C01179 V=7.0 ACC=20 DEC=20
MOVL C01180 V=7.0 ACC=20 DEC=20
ARCOF
TIMER T=30
MOVL C01181 V=11.0 ACC=20 DEC=20
*LAG10
MACRO1 MJ#(0) ARGF2
ARCON
MOVL C01182 V=7.0 ACC=20 DEC=20
MOVL C01183 V=7.0 ACC=20 DEC=20
MOVL C01184 V=7.0 ACC=20 DEC=20
MOVL C01185 V=7.0 ACC=20 DEC=20
MOVL C01186 V=7.0 ACC=20 DEC=20
MOVL C01187 V=7.0 ACC=20 DEC=20
MOVL C01188 V=7.0 ACC=20 DEC=20
MOVL C01189 V=7.0 ACC=20 DEC=20
MOVL C01190 V=7.0 ACC=20 DEC=20
MOVL C01191 V=7.0 PL=1
MOVL C01192 V=7.0 ACC=20 DEC=20
MOVL C01193 V=7.0 ACC=20 DEC=20
MOVL C01194 V=7.0 ACC=20 DEC=20
MOVL C01195 V=7.0 ACC=20 DEC=20
MOVL C01196 V=7.0 ACC=20 DEC=20
MOVL C01197 V=7.0 ACC=20 DEC=20
MOVL C01198 V=7.0 ACC=20 DEC=20
MOVL C01199 V=7.0 ACC=20 DEC=20
MOVL C01200 V=7.0 ACC=20 DEC=20
MOVL C01201 V=7.0 ACC=20 DEC=20
MOVL C01202 V=7.0 ACC=20 DEC=20
MOVL C01203 V=7.0 ACC=20 DEC=20
MOVL C01204 V=7.0 ACC=20 DEC=20
MOVL C01205 V=7.0 ACC=20 DEC=20
MOVL C01206 V=7.0 ACC=20 DEC=20
MOVL C01207 V=7.0 ACC=20 DEC=20
MOVL C01208 V=7.0 ACC=20 DEC=20
MOVL C01209 V=7.0 ACC=20 DEC=20
MOVL C01210 V=7.0 ACC=20 DEC=20
MOVL C01211 V=7.0 ACC=20 DEC=20
MOVL C01212 V=7.0 ACC=20 DEC=20
MOVL C01213 V=7.0 PL=1
MOVL C01214 V=7.0 ACC=20 DEC=20
MOVL C01215 V=7.0 ACC=20 DEC=20
MOVL C01216 V=7.0 ACC=20 DEC=20
MOVL C01217 V=7.0 ACC=20 DEC=20
MOVL C01218 V=7.0 ACC=20 DEC=20
MOVL C01219 V=7.0 ACC=20 DEC=20
MOVL C01220 V=7.0 ACC=20 DEC=20
MOVL C01221 V=7.0 ACC=20 DEC=20
MOVL C01222 V=7.0 ACC=20 DEC=20
MOVC C01223 V=12.0 ACC=20 DEC=20
MOVC C01224 V=12.0 ACC=20 DEC=20
MOVC C01225 V=12.0 ACC=20 DEC=20
MOVL C01226 V=7.0 ACC=20 DEC=20
MOVL C01227 V=7.0 ACC=20 DEC=20
MOVL C01228 V=7.0 ACC=20 DEC=20
MOVL C01229 V=7.0 ACC=20 DEC=20
MOVL C01230 V=7.0 ACC=20 DEC=20
MOVL C01231 V=7.0 ACC=20 DEC=20
MOVL C01232 V=7.0 ACC=20 DEC=20
MOVL C01233 V=7.0 ACC=20 DEC=20
MOVL C01234 V=7.0 ACC=20 DEC=20
MOVL C01235 V=7.0 ACC=20 DEC=20
MOVL C01236 V=7.0 ACC=20 DEC=20
MOVL C01237 V=7.0 ACC=20 DEC=20
MOVL C01238 V=7.0 ACC=20 DEC=20
MOVL C01239 V=7.0 ACC=20 DEC=20
MOVL C01240 V=7.0 ACC=20 DEC=20
MOVL C01241 V=7.0 ACC=20 DEC=20
MOVL C01242 V=7.0 ACC=20 DEC=20
MOVL C01243 V=7.0 ACC=20 DEC=20
MOVL C01244 V=7.0 ACC=20 DEC=20
MOVC C01245 V=12.0 ACC=20 DEC=20
MOVC C01246 V=12.0 ACC=20 DEC=20
MOVC C01247 V=12.0 ACC=20 DEC=20
MOVL C01248 V=7.0 ACC=20 DEC=20
MOVL C01249 V=7.0 ACC=20 DEC=20
MOVL C01250 V=7.0 ACC=20 DEC=20
MOVL C01251 V=7.0 ACC=20 DEC=20
MOVL C01252 V=7.0 ACC=20 DEC=20
MOVL C01253 V=7.0 ACC=20 DEC=20
MOVL C01254 V=7.0 ACC=20 DEC=20
MOVL C01255 V=7.0 ACC=20 DEC=20
MOVL C01256 V=7.0 ACC=20 DEC=20
MOVL C01257 V=7.0 PL=1
MOVL C01258 V=7.0 ACC=20 DEC=20
MOVL C01259 V=7.0 ACC=20 DEC=20
MOVL C01260 V=7.0 ACC=20 DEC=20
MOVL C01261 V=7.0 ACC=20 DEC=20
MOVL C01262 V=7.0 ACC=20 DEC=20
MOVL C01263 V=7.0 ACC=20 DEC=20
MOVL C01264 V=7.0 ACC=20 DEC=20
MOVL C01265 V=7.0 ACC=20 DEC=20
MOVL C01266 V=7.0 ACC=20 DEC=20
MOVL C01267 V=7.0 ACC=20 DEC=20
MOVL C01268 V=7.0 ACC=20 DEC=20
MOVL C01269 V=7.0 ACC=20 DEC=20
MOVL C01270 V=7.0 ACC=20 DEC=20
MOVL C01271 V=7.0 ACC=20 DEC=20
MOVL C01272 V=7.0 ACC=20 DEC=20
MOVL C01273 V=7.0 ACC=20 DEC=20
MOVL C01274 V=7.0 ACC=20 DEC=20
MOVL C01275 V=7.0 ACC=20 DEC=20
MOVL C01276 V=7.0 ACC=20 DEC=20
MOVL C01277 V=7.0 ACC=20 DEC=20
MOVL C01278 V=7.0 ACC=20 DEC=20
MOVL C01279 V=7.0 PL=1
MOVL C01280 V=7.0 ACC=20 DEC=20
MOVL C01281 V=7.0 ACC=20 DEC=20
MOVL C01282 V=7.0 ACC=20 DEC=20
MOVL C01283 V=7.0 ACC=20 DEC=20
MOVL C01284 V=7.0 ACC=20 DEC=20
MOVL C01285 V=7.0 ACC=20 DEC=20
MOVL C01286 V=7.0 ACC=20 DEC=20
MOVL C01287 V=7.0 ACC=20 DEC=20
MOVL C01288 V=7.0 ACC=20 DEC=20
MOVC C01289 V=12.0 ACC=20 DEC=20
MOVC C01290 V=12.0 ACC=20 DEC=20
MOVC C01291 V=12.0 ACC=20 DEC=20
MOVL C01292 V=7.0 ACC=20 DEC=20
MOVL C01293 V=7.0 ACC=20 DEC=20
MOVL C01294 V=7.0 ACC=20 DEC=20
MOVL C01295 V=7.0 ACC=20 DEC=20
MOVL C01296 V=7.0 ACC=20 DEC=20
MOVL C01297 V=7.0 ACC=20 DEC=20
MOVL C01298 V=7.0 ACC=20 DEC=20
MOVL C01299 V=7.0 ACC=20 DEC=20
MOVL C01300 V=7.0 ACC=20 DEC=20
MOVL C01301 V=7.0 ACC=20 DEC=20
MOVL C01302 V=7.0 ACC=20 DEC=20
MOVL C01303 V=7.0 ACC=20 DEC=20
MOVL C01304 V=7.0 ACC=20 DEC=20
MOVL C01305 V=7.0 ACC=20 DEC=20
MOVL C01306 V=7.0 ACC=20 DEC=20
MOVL C01307 V=7.0 ACC=20 DEC=20
MOVL C01308 V=7.0 ACC=20 DEC=20
MOVL C01309 V=7.0 ACC=20 DEC=20
MOVL C01310 V=7.0 ACC=20 DEC=20
MOVL C01311 V=7.0 ACC=20 DEC=20
ARCOF
TIMER T=30
MOVL C01312 V=11.0 ACC=20 DEC=20
*LAG11
MACRO1 MJ#(0) ARGF2
ARCON
MOVL C01313 V=7.0 ACC=20 DEC=20
MOVL C01314 V=7.0 ACC=20 DEC=20
MOVL C01315 V=7.0 ACC=20 DEC=20
MOVL C01316 V=7.0 ACC=20 DEC=20
MOVL C01317 V=7.0 ACC=20 DEC=20
MOVL C01318 V=7.0 ACC=20 DEC=20
MOVL C01319 V=7.0 ACC=20 DEC=20
MOVL C01320 V=7.0 ACC=20 DEC=20
MOVL C01321 V=7.0 ACC=20 DEC=20
MOVL C01322 V=7.0 ACC=20 DEC=20
MOVL C01323 V=7.0 ACC=20 DEC=20
MOVL C01324 V=7.0 ACC=20 DEC=20
MOVL C01325 V=7.0 ACC=20 DEC=20
MOVL C01326 V=7.0 ACC=20 DEC=20
MOVL C01327 V=7.0 ACC=20 DEC=20
MOVL C01328 V=7.0 ACC=20 DEC=20
MOVL C01329 V=7.0 ACC=20 DEC=20
MOVL C01330 V=7.0 ACC=20 DEC=20
MOVL C01331 V=7.0 ACC=20 DEC=20
MOVC C01332 V=12.0 ACC=20 DEC=20
MOVC C01333 V=12.0 ACC=20 DEC=20
MOVC C01334 V=12.0 ACC=20 DEC=20
MOVL C01335 V=7.0 ACC=20 DEC=20
MOVL C01336 V=7.0 ACC=20 DEC=20
MOVL C01337 V=7.0 ACC=20 DEC=20
MOVL C01338 V=7.0 ACC=20 DEC=20
MOVL C01339 V=7.0 ACC=20 DEC=20
MOVL C01340 V=7.0 ACC=20 DEC=20
MOVL C01341 V=7.0 ACC=20 DEC=20
MOVL C01342 V=7.0 ACC=20 DEC=20
MOVL C01343 V=7.0 ACC=20 DEC=20
MOVL C01344 V=7.0 PL=1
MOVL C01345 V=7.0 ACC=20 DEC=20
MOVL C01346 V=7.0 ACC=20 DEC=20
MOVL C01347 V=7.0 ACC=20 DEC=20
MOVL C01348 V=7.0 ACC=20 DEC=20
MOVL C01349 V=7.0 ACC=20 DEC=20
MOVL C01350 V=7.0 ACC=20 DEC=20
MOVL C01351 V=7.0 ACC=20 DEC=20
MOVL C01352 V=7.0 ACC=20 DEC=20
MOVL C01353 V=7.0 ACC=20 DEC=20
MOVL C01354 V=7.0 ACC=20 DEC=20
MOVL C01355 V=7.0 ACC=20 DEC=20
MOVL C01356 V=7.0 ACC=20 DEC=20
MOVL C01357 V=7.0 ACC=20 DEC=20
MOVL C01358 V=7.0 ACC=20 DEC=20
MOVL C01359 V=7.0 ACC=20 DEC=20
MOVL C01360 V=7.0 ACC=20 DEC=20
MOVL C01361 V=7.0 ACC=20 DEC=20
MOVL C01362 V=7.0 ACC=20 DEC=20
MOVL C01363 V=7.0 ACC=20 DEC=20
MOVL C01364 V=7.0 ACC=20 DEC=20
MOVL C01365 V=7.0 ACC=20 DEC=20
MOVL C01366 V=7.0 PL=1
MOVL C01367 V=7.0 ACC=20 DEC=20
MOVL C01368 V=7.0 ACC=20 DEC=20
MOVL C01369 V=7.0 ACC=20 DEC=20
MOVL C01370 V=7.0 ACC=20 DEC=20
MOVL C01371 V=7.0 ACC=20 DEC=20
MOVL C01372 V=7.0 ACC=20 DEC=20
MOVL C01373 V=7.0 ACC=20 DEC=20
MOVL C01374 V=7.0 ACC=20 DEC=20
MOVL C01375 V=7.0 ACC=20 DEC=20
MOVC C01376 V=12.0 ACC=20 DEC=20
MOVC C01377 V=12.0 ACC=20 DEC=20
MOVC C01378 V=12.0 ACC=20 DEC=20
MOVL C01379 V=7.0 ACC=20 DEC=20
MOVL C01380 V=7.0 ACC=20 DEC=20
MOVL C01381 V=7.0 ACC=20 DEC=20
MOVL C01382 V=7.0 ACC=20 DEC=20
MOVL C01383 V=7.0 ACC=20 DEC=20
MOVL C01384 V=7.0 ACC=20 DEC=20
MOVL C01385 V=7.0 ACC=20 DEC=20
MOVL C01386 V=7.0 ACC=20 DEC=20
MOVL C01387 V=7.0 ACC=20 DEC=20
MOVL C01388 V=7.0 ACC=20 DEC=20
MOVL C01389 V=7.0 ACC=20 DEC=20
MOVL C01390 V=7.0 ACC=20 DEC=20
MOVL C01391 V=7.0 ACC=20 DEC=20
MOVL C01392 V=7.0 ACC=20 DEC=20
MOVL C01393 V=7.0 ACC=20 DEC=20
MOVL C01394 V=7.0 ACC=20 DEC=20
MOVL C01395 V=7.0 ACC=20 DEC=20
MOVL C01396 V=7.0 ACC=20 DEC=20
MOVL C01397 V=7.0 ACC=20 DEC=20
MOVC C01398 V=12.0 ACC=20 DEC=20
MOVC C01399 V=12.0 ACC=20 DEC=20
MOVC C01400 V=12.0 ACC=20 DEC=20
MOVL C01401 V=7.0 ACC=20 DEC=20
MOVL C01402 V=7.0 ACC=20 DEC=20
MOVL C01403 V=7.0 ACC=20 DEC=20
MOVL C01404 V=7.0 ACC=20 DEC=20
MOVL C01405 V=7.0 ACC=20 DEC=20
MOVL C01406 V=7.0 ACC=20 DEC=20
MOVL C01407 V=7.0 ACC=20 DEC=20
MOVL C01408 V=7.0 ACC=20 DEC=20
MOVL C01409 V=7.0 ACC=20 DEC=20
MOVL C01410 V=7.0 PL=1
MOVL C01411 V=7.0 ACC=20 DEC=20
MOVL C01412 V=7.0 ACC=20 DEC=20
MOVL C01413 V=7.0 ACC=20 DEC=20
MOVL C01414 V=7.0 ACC=20 DEC=20
MOVL C01415 V=7.0 ACC=20 DEC=20
MOVL C01416 V=7.0 ACC=20 DEC=20
MOVL C01417 V=7.0 ACC=20 DEC=20
MOVL C01418 V=7.0 ACC=20 DEC=20
MOVL C01419 V=7.0 ACC=20 DEC=20
MOVL C01420 V=7.0 ACC=20 DEC=20
MOVL C01421 V=7.0 ACC=20 DEC=20
MOVL C01422 V=7.0 ACC=20 DEC=20
MOVL C01423 V=7.0 ACC=20 DEC=20
MOVL C01424 V=7.0 ACC=20 DEC=20
MOVL C01425 V=7.0 ACC=20 DEC=20
MOVL C01426 V=7.0 ACC=20 DEC=20
MOVL C01427 V=7.0 ACC=20 DEC=20
MOVL C01428 V=7.0 ACC=20 DEC=20
MOVL C01429 V=7.0 ACC=20 DEC=20
MOVL C01430 V=7.0 ACC=20 DEC=20
MOVL C01431 V=7.0 ACC=20 DEC=20
MOVL C01432 V=7.0 PL=1
MOVL C01433 V=7.0 ACC=20 DEC=20
MOVL C01434 V=7.0 ACC=20 DEC=20
MOVL C01435 V=7.0 ACC=20 DEC=20
MOVL C01436 V=7.0 ACC=20 DEC=20
MOVL C01437 V=7.0 ACC=20 DEC=20
MOVL C01438 V=7.0 ACC=20 DEC=20
MOVL C01439 V=7.0 ACC=20 DEC=20
MOVL C01440 V=7.0 ACC=20 DEC=20
MOVL C01441 V=7.0 ACC=20 DEC=20
MOVL C01442 V=7.0 ACC=20 DEC=20
ARCOF
TIMER T=30
MOVL C01443 V=11.0 ACC=20 DEC=20
*LAG12
MACRO1 MJ#(0) ARGF2
ARCON
MOVL C01444 V=7.0 ACC=20 DEC=20
MOVL C01445 V=7.0 ACC=20 DEC=20
MOVL C01446 V=7.0 ACC=20 DEC=20
MOVL C01447 V=7.0 ACC=20 DEC=20
MOVL C01448 V=7.0 ACC=20 DEC=20
MOVL C01449 V=7.0 ACC=20 DEC=20
MOVL C01450 V=7.0 ACC=20 DEC=20
MOVL C01451 V=7.0 ACC=20 DEC=20
MOVL C01452 V=7.0 ACC=20 DEC=20
MOVL C01453 V=7.0 PL=1
MOVL C01454 V=7.0 ACC=20 DEC=20
MOVL C01455 V=7.0 ACC=20 DEC=20
MOVL C01456 V=7.0 ACC=20 DEC=20
MOVL C01457 V=7.0 ACC=20 DEC=20
MOVL C01458 V=7.0 ACC=20 DEC=20
MOVL C01459 V=7.0 ACC=20 DEC=20
MOVL C01460 V=7.0 ACC=20 DEC=20
MOVL C01461 V=7.0 ACC=20 DEC=20
MOVL C01462 V=7.0 ACC=20 DEC=20
MOVL C01463 V=7.0 ACC=20 DEC=20
MOVL C01464 V=7.0 ACC=20 DEC=20
MOVL C01465 V=7.0 ACC=20 DEC=20
MOVL C01466 V=7.0 ACC=20 DEC=20
MOVL C01467 V=7.0 ACC=20 DEC=20
MOVL C01468 V=7.0 ACC=20 DEC=20
MOVL C01469 V=7.0 ACC=20 DEC=20
MOVL C01470 V=7.0 ACC=20 DEC=20
MOVL C01471 V=7.0 ACC=20 DEC=20
MOVL C01472 V=7.0 ACC=20 DEC=20
MOVL C01473 V=7.0 ACC=20 DEC=20
MOVL C01474 V=7.0 ACC=20 DEC=20
MOVL C01475 V=7.0 PL=1
MOVL C01476 V=7.0 ACC=20 DEC=20
MOVL C01477 V=7.0 ACC=20 DEC=20
MOVL C01478 V=7.0 ACC=20 DEC=20
MOVL C01479 V=7.0 ACC=20 DEC=20
MOVL C01480 V=7.0 ACC=20 DEC=20
MOVL C01481 V=7.0 ACC=20 DEC=20
MOVL C01482 V=7.0 ACC=20 DEC=20
MOVL C01483 V=7.0 ACC=20 DEC=20
MOVL C01484 V=7.0 ACC=20 DEC=20
MOVC C01485 V=12.0 ACC=20 DEC=20
MOVC C01486 V=12.0 ACC=20 DEC=20
MOVC C01487 V=12.0 ACC=20 DEC=20
MOVL C01488 V=7.0 ACC=20 DEC=20
MOVL C01489 V=7.0 ACC=20 DEC=20
MOVL C01490 V=7.0 ACC=20 DEC=20
MOVL C01491 V=7.0 ACC=20 DEC=20
MOVL C01492 V=7.0 ACC=20 DEC=20
MOVL C01493 V=7.0 ACC=20 DEC=20
MOVL C01494 V=7.0 ACC=20 DEC=20
MOVL C01495 V=7.0 ACC=20 DEC=20
MOVL C01496 V=7.0 ACC=20 DEC=20
MOVL C01497 V=7.0 ACC=20 DEC=20
MOVL C01498 V=7.0 ACC=20 DEC=20
MOVL C01499 V=7.0 ACC=20 DEC=20
MOVL C01500 V=7.0 ACC=20 DEC=20
MOVL C01501 V=7.0 ACC=20 DEC=20
MOVL C01502 V=7.0 ACC=20 DEC=20
MOVL C01503 V=7.0 ACC=20 DEC=20
MOVL C01504 V=7.0 ACC=20 DEC=20
MOVL C01505 V=7.0 ACC=20 DEC=20
MOVL C01506 V=7.0 ACC=20 DEC=20
MOVC C01507 V=12.0 ACC=20 DEC=20
MOVC C01508 V=12.0 ACC=20 DEC=20
MOVC C01509 V=12.0 ACC=20 DEC=20
MOVL C01510 V=7.0 ACC=20 DEC=20
MOVL C01511 V=7.0 ACC=20 DEC=20
MOVL C01512 V=7.0 ACC=20 DEC=20
MOVL C01513 V=7.0 ACC=20 DEC=20
MOVL C01514 V=7.0 ACC=20 DEC=20
MOVL C01515 V=7.0 ACC=20 DEC=20
MOVL C01516 V=7.0 ACC=20 DEC=20
MOVL C01517 V=7.0 ACC=20 DEC=20
MOVL C01518 V=7.0 ACC=20 DEC=20
MOVL C01519 V=7.0 PL=1
MOVL C01520 V=7.0 ACC=20 DEC=20
MOVL C01521 V=7.0 ACC=20 DEC=20
MOVL C01522 V=7.0 ACC=20 DEC=20
MOVL C01523 V=7.0 ACC=20 DEC=20
MOVL C01524 V=7.0 ACC=20 DEC=20
MOVL C01525 V=7.0 ACC=20 DEC=20
MOVL C01526 V=7.0 ACC=20 DEC=20
MOVL C01527 V=7.0 ACC=20 DEC=20
MOVL C01528 V=7.0 ACC=20 DEC=20
MOVL C01529 V=7.0 ACC=20 DEC=20
MOVL C01530 V=7.0 ACC=20 DEC=20
MOVL C01531 V=7.0 ACC=20 DEC=20
MOVL C01532 V=7.0 ACC=20 DEC=20
MOVL C01533 V=7.0 ACC=20 DEC=20
MOVL C01534 V=7.0 ACC=20 DEC=20
MOVL C01535 V=7.0 ACC=20 DEC=20
MOVL C01536 V=7.0 ACC=20 DEC=20
MOVL C01537 V=7.0 ACC=20 DEC=20
MOVL C01538 V=7.0 ACC=20 DEC=20
MOVL C01539 V=7.0 ACC=20 DEC=20
MOVL C01540 V=7.0 ACC=20 DEC=20
MOVL C01541 V=7.0 PL=1
MOVL C01542 V=7.0 ACC=20 DEC=20
MOVL C01543 V=7.0 ACC=20 DEC=20
MOVL C01544 V=7.0 ACC=20 DEC=20
MOVL C01545 V=7.0 ACC=20 DEC=20
MOVL C01546 V=7.0 ACC=20 DEC=20
MOVL C01547 V=7.0 ACC=20 DEC=20
MOVL C01548 V=7.0 ACC=20 DEC=20
MOVL C01549 V=7.0 ACC=20 DEC=20
MOVL C01550 V=7.0 ACC=20 DEC=20
MOVC C01551 V=12.0 ACC=20 DEC=20
MOVC C01552 V=12.0 ACC=20 DEC=20
MOVC C01553 V=12.0 ACC=20 DEC=20
MOVL C01554 V=7.0 ACC=20 DEC=20
MOVL C01555 V=7.0 ACC=20 DEC=20
MOVL C01556 V=7.0 ACC=20 DEC=20
MOVL C01557 V=7.0 ACC=20 DEC=20
MOVL C01558 V=7.0 ACC=20 DEC=20
MOVL C01559 V=7.0 ACC=20 DEC=20
MOVL C01560 V=7.0 ACC=20 DEC=20
MOVL C01561 V=7.0 ACC=20 DEC=20
MOVL C01562 V=7.0 ACC=20 DEC=20
MOVL C01563 V=7.0 ACC=20 DEC=20
MOVL C01564 V=7.0 ACC=20 DEC=20
MOVL C01565 V=7.0 ACC=20 DEC=20
MOVL C01566 V=7.0 ACC=20 DEC=20
MOVL C01567 V=7.0 ACC=20 DEC=20
MOVL C01568 V=7.0 ACC=20 DEC=20
MOVL C01569 V=7.0 ACC=20 DEC=20
MOVL C01570 V=7.0 ACC=20 DEC=20
MOVL C01571 V=7.0 ACC=20 DEC=20
MOVL C01572 V=7.0 ACC=20 DEC=20
MOVL C01573 V=7.0 ACC=20 DEC=20
ARCOF
TIMER T=30
MOVL C01574 V=11.0 ACC=20 DEC=20
*LAG13
MACRO1 MJ#(0) ARGF2
ARCON
MOVL C01575 V=7.0 ACC=20 DEC=20
MOVL C01576 V=7.0 ACC=20 DEC=20
MOVL C01577 V=7.0 ACC=20 DEC=20
MOVL C01578 V=7.0 ACC=20 DEC=20
MOVL C01579 V=7.0 ACC=20 DEC=20
MOVL C01580 V=7.0 ACC=20 DEC=20
MOVL C01581 V=7.0 ACC=20 DEC=20
MOVL C01582 V=7.0 ACC=20 DEC=20
MOVL C01583 V=7.0 ACC=20 DEC=20
MOVL C01584 V=7.0 ACC=20 DEC=20
MOVL C01585 V=7.0 ACC=20 DEC=20
MOVL C01586 V=7.0 ACC=20 DEC=20
MOVL C01587 V=7.0 ACC=20 DEC=20
MOVL C01588 V=7.0 ACC=20 DEC=20
MOVL C01589 V=7.0 ACC=20 DEC=20
MOVL C01590 V=7.0 ACC=20 DEC=20
MOVL C01591 V=7.0 ACC=20 DEC=20
MOVL C01592 V=7.0 ACC=20 DEC=20
MOVL C01593 V=7.0 ACC=20 DEC=20
MOVC C01594 V=12.0 ACC=20 DEC=20
MOVC C01595 V=12.0 ACC=20 DEC=20
MOVC C01596 V=12.0 ACC=20 DEC=20
MOVL C01597 V=7.0 ACC=20 DEC=20
MOVL C01598 V=7.0 ACC=20 DEC=20
MOVL C01599 V=7.0 ACC=20 DEC=20
MOVL C01600 V=7.0 ACC=20 DEC=20
MOVL C01601 V=7.0 ACC=20 DEC=20
MOVL C01602 V=7.0 ACC=20 DEC=20
MOVL C01603 V=7.0 ACC=20 DEC=20
MOVL C01604 V=7.0 ACC=20 DEC=20
MOVL C01605 V=7.0 ACC=20 DEC=20
MOVL C01606 V=7.0 PL=1
MOVL C01607 V=7.0 ACC=20 DEC=20
MOVL C01608 V=7.0 ACC=20 DEC=20
MOVL C01609 V=7.0 ACC=20 DEC=20
MOVL C01610 V=7.0 ACC=20 DEC=20
MOVL C01611 V=7.0 ACC=20 DEC=20
MOVL C01612 V=7.0 ACC=20 DEC=20
MOVL C01613 V=7.0 ACC=20 DEC=20
MOVL C01614 V=7.0 ACC=20 DEC=20
MOVL C01615 V=7.0 ACC=20 DEC=20
MOVL C01616 V=7.0 ACC=20 DEC=20
MOVL C01617 V=7.0 ACC=20 DEC=20
MOVL C01618 V=7.0 ACC=20 DEC=20
MOVL C01619 V=7.0 ACC=20 DEC=20
MOVL C01620 V=7.0 ACC=20 DEC=20
MOVL C01621 V=7.0 ACC=20 DEC=20
MOVL C01622 V=7.0 ACC=20 DEC=20
MOVL C01623 V=7.0 ACC=20 DEC=20
MOVL C01624 V=7.0 ACC=20 DEC=20
MOVL C01625 V=7.0 ACC=20 DEC=20
MOVL C01626 V=7.0 ACC=20 DEC=20
MOVL C01627 V=7.0 ACC=20 DEC=20
MOVL C01628 V=7.0 PL=1
MOVL C01629 V=7.0 ACC=20 DEC=20
MOVL C01630 V=7.0 ACC=20 DEC=20
MOVL C01631 V=7.0 ACC=20 DEC=20
MOVL C01632 V=7.0 ACC=20 DEC=20
MOVL C01633 V=7.0 ACC=20 DEC=20
MOVL C01634 V=7.0 ACC=20 DEC=20
MOVL C01635 V=7.0 ACC=20 DEC=20
MOVL C01636 V=7.0 ACC=20 DEC=20
MOVL C01637 V=7.0 ACC=20 DEC=20
MOVC C01638 V=12.0 ACC=20 DEC=20
MOVC C01639 V=12.0 ACC=20 DEC=20
MOVC C01640 V=12.0 ACC=20 DEC=20
MOVL C01641 V=7.0 ACC=20 DEC=20
MOVL C01642 V=7.0 ACC=20 DEC=20
MOVL C01643 V=7.0 ACC=20 DEC=20
MOVL C01644 V=7.0 ACC=20 DEC=20
MOVL C01645 V=7.0 ACC=20 DEC=20
MOVL C01646 V=7.0 ACC=20 DEC=20
MOVL C01647 V=7.0 ACC=20 DEC=20
MOVL C01648 V=7.0 ACC=20 DEC=20
MOVL C01649 V=7.0 ACC=20 DEC=20
MOVL C01650 V=7.0 ACC=20 DEC=20
MOVL C01651 V=7.0 ACC=20 DEC=20
MOVL C01652 V=7.0 ACC=20 DEC=20
MOVL C01653 V=7.0 ACC=20 DEC=20
MOVL C01654 V=7.0 ACC=20 DEC=20
MOVL C01655 V=7.0 ACC=20 DEC=20
MOVL C01656 V=7.0 ACC=20 DEC=20
MOVL C01657 V=7.0 ACC=20 DEC=20
MOVL C01658 V=7.0 ACC=20 DEC=20
MOVL C01659 V=7.0 ACC=20 DEC=20
MOVC C01660 V=12.0 ACC=20 DEC=20
MOVC C01661 V=12.0 ACC=20 DEC=20
MOVC C01662 V=12.0 ACC=20 DEC=20
MOVL C01663 V=7.0 ACC=20 DEC=20
MOVL C01664 V=7.0 ACC=20 DEC=20
MOVL C01665 V=7.0 ACC=20 DEC=20
MOVL C01666 V=7.0 ACC=20 DEC=20
MOVL C01667 V=7.0 ACC=20 DEC=20
MOVL C01668 V=7.0 ACC=20 DEC=20
MOVL C01669 V=7.0 ACC=20 DEC=20
MOVL C01670 V=7.0 ACC=20 DEC=20
MOVL C01671 V=7.0 ACC=20 DEC=20
MOVL C01672 V=7.0 PL=1
MOVL C01673 V=7.0 ACC=20 DEC=20
MOVL C01674 V=7.0 ACC=20 DEC=20
MOVL C01675 V=7.0 ACC=20 DEC=20
MOVL C01676 V=7.0 ACC=20 DEC=20
MOVL C01677 V=7.0 ACC=20 DEC=20
MOVL C01678 V=7.0 ACC=20 DEC=20
MOVL C01679 V=7.0 ACC=20 DEC=20
MOVL C01680 V=7.0 ACC=20 DEC=20
MOVL C01681 V=7.0 ACC=20 DEC=20
MOVL C01682 V=7.0 ACC=20 DEC=20
MOVL C01683 V=7.0 ACC=20 DEC=20
MOVL C01684 V=7.0 ACC=20 DEC=20
MOVL C01685 V=7.0 ACC=20 DEC=20
MOVL C01686 V=7.0 ACC=20 DEC=20
MOVL C01687 V=7.0 ACC=20 DEC=20
MOVL C01688 V=7.0 ACC=20 DEC=20
MOVL C01689 V=7.0 ACC=20 DEC=20
MOVL C01690 V=7.0 ACC=20 DEC=20
MOVL C01691 V=7.0 ACC=20 DEC=20
MOVL C01692 V=7.0 ACC=20 DEC=20
MOVL C01693 V=7.0 ACC=20 DEC=20
MOVL C01694 V=7.0 PL=1
MOVL C01695 V=7.0 ACC=20 DEC=20
MOVL C01696 V=7.0 ACC=20 DEC=20
MOVL C01697 V=7.0 ACC=20 DEC=20
MOVL C01698 V=7.0 ACC=20 DEC=20
MOVL C01699 V=7.0 ACC=20 DEC=20
MOVL C01700 V=7.0 ACC=20 DEC=20
MOVL C01701 V=7.0 ACC=20 DEC=20
MOVL C01702 V=7.0 ACC=20 DEC=20
MOVL C01703 V=7.0 ACC=20 DEC=20
MOVL C01704 V=7.0 ACC=20 DEC=20
ARCOF
TIMER T=30
MOVL C01705 V=11.0 ACC=20 DEC=20
*LAG14
MACRO1 MJ#(0) ARGF2
ARCON
MOVL C01706 V=7.0 ACC=20 DEC=20
MOVL C01707 V=7.0 ACC=20 DEC=20
MOVL C01708 V=7.0 ACC=20 DEC=20
MOVL C01709 V=7.0 ACC=20 DEC=20
MOVL C01710 V=7.0 ACC=20 DEC=20
MOVL C01711 V=7.0 ACC=20 DEC=20
MOVL C01712 V=7.0 ACC=20 DEC=20
MOVL C01713 V=7.0 ACC=20 DEC=20
MOVL C01714 V=7.0 ACC=20 DEC=20
MOVL C01715 V=7.0 PL=1
MOVL C01716 V=7.0 ACC=20 DEC=20
MOVL C01717 V=7.0 ACC=20 DEC=20
MOVL C01718 V=7.0 ACC=20 DEC=20
MOVL C01719 V=7.0 ACC=20 DEC=20
MOVL C01720 V=7.0 ACC=20 DEC=20
MOVL C01721 V=7.0 ACC=20 DEC=20
MOVL C01722 V=7.0 ACC=20 DEC=20
MOVL C01723 V=7.0 ACC=20 DEC=20
MOVL C01724 V=7.0 ACC=20 DEC=20
MOVL C01725 V=7.0 ACC=20 DEC=20
MOVL C01726 V=7.0 ACC=20 DEC=20
MOVL C01727 V=7.0 ACC=20 DEC=20
MOVL C01728 V=7.0 ACC=20 DEC=20
MOVL C01729 V=7.0 ACC=20 DEC=20
MOVL C01730 V=7.0 ACC=20 DEC=20
MOVL C01731 V=7.0 ACC=20 DEC=20
MOVL C01732 V=7.0 ACC=20 DEC=20
MOVL C01733 V=7.0 ACC=20 DEC=20
MOVL C01734 V=7.0 ACC=20 DEC=20
MOVL C01735 V=7.0 ACC=20 DEC=20
MOVL C01736 V=7.0 ACC=20 DEC=20
MOVL C01737 V=7.0 PL=1
MOVL C01738 V=7.0 ACC=20 DEC=20
MOVL C01739 V=7.0 ACC=20 DEC=20
MOVL C01740 V=7.0 ACC=20 DEC=20
MOVL C01741 V=7.0 ACC=20 DEC=20
MOVL C01742 V=7.0 ACC=20 DEC=20
MOVL C01743 V=7.0 ACC=20 DEC=20
MOVL C01744 V=7.0 ACC=20 DEC=20
MOVL C01745 V=7.0 ACC=20 DEC=20
MOVL C01746 V=7.0 ACC=20 DEC=20
MOVC C01747 V=12.0 ACC=20 DEC=20
MOVC C01748 V=12.0 ACC=20 DEC=20
MOVC C01749 V=12.0 ACC=20 DEC=20
MOVL C01750 V=7.0 ACC=20 DEC=20
MOVL C01751 V=7.0 ACC=20 DEC=20
MOVL C01752 V=7.0 ACC=20 DEC=20
MOVL C01753 V=7.0 ACC=20 DEC=20
MOVL C01754 V=7.0 ACC=20 DEC=20
MOVL C01755 V=7.0 ACC=20 DEC=20
MOVL C01756 V=7.0 ACC=20 DEC=20
MOVL C01757 V=7.0 ACC=20 DEC=20
MOVL C01758 V=7.0 ACC=20 DEC=20
MOVL C01759 V=7.0 ACC=20 DEC=20
MOVL C01760 V=7.0 ACC=20 DEC=20
MOVL C01761 V=7.0 ACC=20 DEC=20
MOVL C01762 V=7.0 ACC=20 DEC=20
MOVL C01763 V=7.0 ACC=20 DEC=20
MOVL C01764 V=7.0 ACC=20 DEC=20
MOVL C01765 V=7.0 ACC=20 DEC=20
MOVL C01766 V=7.0 ACC=20 DEC=20
MOVL C01767 V=7.0 ACC=20 DEC=20
MOVL C01768 V=7.0 ACC=20 DEC=20
MOVC C01769 V=12.0 ACC=20 DEC=20
MOVC C01770 V=12.0 ACC=20 DEC=20
MOVC C01771 V=12.0 ACC=20 DEC=20
MOVL C01772 V=7.0 ACC=20 DEC=20
MOVL C01773 V=7.0 ACC=20 DEC=20
MOVL C01774 V=7.0 ACC=20 DEC=20
MOVL C01775 V=7.0 ACC=20 DEC=20
MOVL C01776 V=7.0 ACC=20 DEC=20
MOVL C01777 V=7.0 ACC=20 DEC=20
MOVL C01778 V=7.0 ACC=20 DEC=20
MOVL C01779 V=7.0 ACC=20 DEC=20
MOVL C01780 V=7.0 ACC=20 DEC=20
MOVL C01781 V=7.0 PL=1
MOVL C01782 V=7.0 ACC=20 DEC=20
MOVL C01783 V=7.0 ACC=20 DEC=20
MOVL C01784 V=7.0 ACC=20 DEC=20
MOVL C01785 V=7.0 ACC=20 DEC=20
MOVL C01786 V=7.0 ACC=20 DEC=20
MOVL C01787 V=7.0 ACC=20 DEC=20
MOVL C01788 V=7.0 ACC=20 DEC=20
MOVL C01789 V=7.0 ACC=20 DEC=20
MOVL C01790 V=7.0 ACC=20 DEC=20
MOVL C01791 V=7.0 ACC=20 DEC=20
MOVL C01792 V=7.0 ACC=20 DEC=20
MOVL C01793 V=7.0 ACC=20 DEC=20
MOVL C01794 V=7.0 ACC=20 DEC=20
MOVL C01795 V=7.0 ACC=20 DEC=20
MOVL C01796 V=7.0 ACC=20 DEC=20
MOVL C01797 V=7.0 ACC=20 DEC=20
MOVL C01798 V=7.0 ACC=20 DEC=20
MOVL C01799 V=7.0 ACC=20 DEC=20
MOVL C01800 V=7.0 ACC=20 DEC=20
MOVL C01801 V=7.0 ACC=20 DEC=20
MOVL C01802 V=7.0 ACC=20 DEC=20
MOVL C01803 V=7.0 PL=1
MOVL C01804 V=7.0 ACC=20 DEC=20
MOVL C01805 V=7.0 ACC=20 DEC=20
MOVL C01806 V=7.0 ACC=20 DEC=20
MOVL C01807 V=7.0 ACC=20 DEC=20
MOVL C01808 V=7.0 ACC=20 DEC=20
MOVL C01809 V=7.0 ACC=20 DEC=20
MOVL C01810 V=7.0 ACC=20 DEC=20
MOVL C01811 V=7.0 ACC=20 DEC=20
MOVL C01812 V=7.0 ACC=20 DEC=20
MOVC C01813 V=12.0 ACC=20 DEC=20
MOVC C01814 V=12.0 ACC=20 DEC=20
MOVC C01815 V=12.0 ACC=20 DEC=20
MOVL C01816 V=7.0 ACC=20 DEC=20
MOVL C01817 V=7.0 ACC=20 DEC=20
MOVL C01818 V=7.0 ACC=20 DEC=20
MOVL C01819 V=7.0 ACC=20 DEC=20
MOVL C01820 V=7.0 ACC=20 DEC=20
MOVL C01821 V=7.0 ACC=20 DEC=20
MOVL C01822 V=7.0 ACC=20 DEC=20
MOVL C01823 V=7.0 ACC=20 DEC=20
MOVL C01824 V=7.0 ACC=20 DEC=20
MOVL C01825 V=7.0 ACC=20 DEC=20
MOVL C01826 V=7.0 ACC=20 DEC=20
MOVL C01827 V=7.0 ACC=20 DEC=20
MOVL C01828 V=7.0 ACC=20 DEC=20
MOVL C01829 V=7.0 ACC=20 DEC=20
MOVL C01830 V=7.0 ACC=20 DEC=20
MOVL C01831 V=7.0 ACC=20 DEC=20
MOVL C01832 V=7.0 ACC=20 DEC=20
MOVL C01833 V=7.0 ACC=20 DEC=20
MOVL C01834 V=7.0 ACC=20 DEC=20
MOVL C01835 V=7.0 ACC=20 DEC=20
ARCOF
TIMER T=30
MOVL C01836 V=11.0 ACC=20 DEC=20
*LAG15
MACRO1 MJ#(0) ARGF2
ARCON
MOVL C01837 V=7.0 ACC=20 DEC=20
MOVL C01838 V=7.0 ACC=20 DEC=20
MOVL C01839 V=7.0 ACC=20 DEC=20
MOVL C01840 V=7.0 ACC=20 DEC=20
MOVL C01841 V=7.0 ACC=20 DEC=20
MOVL C01842 V=7.0 ACC=20 DEC=20
MOVL C01843 V=7.0 ACC=20 DEC=20
MOVL C01844 V=7.0 ACC=20 DEC=20
MOVL C01845 V=7.0 ACC=20 DEC=20
MOVL C01846 V=7.0 ACC=20 DEC=20
MOVL C01847 V=7.0 ACC=20 DEC=20
MOVL C01848 V=7.0 ACC=20 DEC=20
MOVL C01849 V=7.0 ACC=20 DEC=20
MOVL C01850 V=7.0 ACC=20 DEC=20
MOVL C01851 V=7.0 ACC=20 DEC=20
MOVL C01852 V=7.0 ACC=20 DEC=20
MOVL C01853 V=7.0 ACC=20 DEC=20
MOVL C01854 V=7.0 ACC=20 DEC=20
MOVL C01855 V=7.0 ACC=20 DEC=20
